(* IEC 61131-3 sources: daoli-st-library/DL_Device (part 27) *)

(* ---- FB_DL_OvenCureProfileSeq.st ---- *)
(*
  Name: FB_DL_OvenCureProfileSeq
  Category: DL_Device
  Version: 1.0.0
  Round: R89 / 2026-11-25
  开源溯源：clean-room 自研（族 涂装喷涂线，ST 开源生态实测 0 命中，无外部代码引入）
  功能：烘干炉固化温度曲线执行顺序：升温→保温→冷却→出炉许可，每段结束判据独立。
  边界条件：① 温度与速率入参全部过非有限闸（含三元素设定数组逐项），配置越域即锁故障（101）；
            ② 保温段使用独立 TON（tonSoak，PT := tSoakS），与升温/冷却段判据不同源，无双窗配比问题（R100）；
            ③ 超温判据以段 1 设定 + 15 ℃ 为上限（固化段为最高温段），越限立即锁故障（102）；
            ④ 出炉许可为单拍脉冲（内部 _bDone 置位 → 出口映射），后驻留 eDone 至启动释放；
            ⑤ 故障解除唯一路径：故障相内 xStart 释放（R152），清锁存回 eIdle。
  状态机：eIdle / eSeg1 / eSeg2 / eSeg3 / eDone / eFault（CASE 含 ELSE 兜底）。
*)
TYPE E_DL_OcpPhase :
(
    eIdle := 0,         (* 待机：等启动沿 / Idle, waiting for start edge *)
    eSeg1 := 10,        (* 段 1 升温：升到固化温度带 / Segment 1, ramp to cure band *)
    eSeg2 := 20,        (* 段 2 保温：保温窗且带内 / Segment 2, soak window in band *)
    eSeg3 := 30,        (* 段 3 冷却：冷到出炉温度 / Segment 3, cool down *)
    eDone := 40,        (* 完成相：出炉许可后驻留 / Done, holds after discharge permit *)
    eFault := 90        (* 故障相：锁存待释放 / Fault latched, awaiting release *)
);
END_TYPE

FUNCTION_BLOCK FB_DL_OvenCureProfileSeq
VAR_INPUT
    xStart : BOOL;                          (* 启动命令（上升沿起序） [-] Start command, rising edge *)
    fTempActC : REAL;                       (* 炉温实测 [℃] Oven temperature actual [degC] *)
    fTempSpC : ARRAY[1..3] OF REAL;         (* 三段温度设定（升温/保温/冷却） [℃] Segment setpoints [degC] *)
    fRampCpm : REAL;                        (* 允许升温速率 [℃/min] Allowed ramp rate [degC/min] *)
    tSoakS : TIME;                          (* 保温窗 [ms] Soak window [ms] *)
    fCoolToC : REAL;                        (* 冷却目标（出炉温度） [℃] Cool-down target [degC] *)
END_VAR
VAR_OUTPUT
    eState : E_DL_OcpPhase;                 (* 当前相 [-] Present phase *)
    nSegIdx : INT;                          (* 当前段号（0 空闲，1~3） [段] Present segment index *)
    xDone : BOOL;                           (* 出炉许可单拍脉冲 [-] Discharge permit pulse *)
    xFault : BOOL;                          (* 故障锁存标志 [-] Fault latched *)
END_VAR
VAR
    _eState : E_DL_OcpPhase := E_DL_OcpPhase.eIdle;  (* 内部相（CASE 唯一写入目标） [-] Internal phase *)
    _bDone : BOOL := FALSE;         (* 单拍完成标志（段 1 预清） [-] One-scan done flag *)
    _bFaultLatch : BOOL := FALSE;   (* 故障锁存位 [-] Fault latch *)
    _bReqFault : BOOL := FALSE;     (* 单拍故障请求（段 1 预清） [-] Fault request *)
    _bCfgBad : BOOL := FALSE;       (* 配置非法当拍量 [-] Configuration bad *)
    _nSeg : INT := 0;               (* 段号保持量 [段] Segment index hold *)
    _nErr : INT := 0;               (* 故障码锁存（101 组态 / 102 超温 / 103 非法相） [-] Latched code *)
    _nReqErr : INT := 0;            (* 当拍请求码 [-] Requested code *)
    _nI : INT := 1;                 (* 设定数组遍历索引 [-] Setpoint loop index *)
    tonSoak : TON;                  (* 保温窗（段 0 无条件调用） / Soak window timer *)
    rtStart : R_TRIG;               (* 启动沿（段 0 无条件调用） / Start edge *)
END_VAR
VAR CONSTANT
    DL_OCP_TOL : REAL := 5.0;           (* 段到位带半宽 [℃] Segment in-band half-width [degC] *)
    DL_OCP_OVER : REAL := 15.0;         (* 超温裕度 [℃] Over-temperature margin [degC] *)
    DL_OCP_T_MIN : REAL := 0.0;         (* 温度下限 [℃] Temperature floor [degC] *)
    DL_OCP_T_MAX : REAL := 400.0;       (* 温度上限 [℃] Temperature ceiling [degC] *)
    DL_OCP_R_MIN : REAL := 0.5;         (* 允许速率下限 [℃/min] Ramp rate floor [degC/min] *)
    DL_OCP_R_MAX : REAL := 50.0;        (* 允许速率上限 [℃/min] Ramp rate ceiling [degC/min] *)
    DL_OCP_SEGN : INT := 3;             (* 设定段数 [-] Segment count *)
END_VAR
(* —— 段 0：沿与保温 TON 无条件周期刷新（R7） —— *)
rtStart(CLK := xStart);                                             (* 启动沿 / Start edge *)
tonSoak(IN := (_eState = E_DL_OcpPhase.eSeg2), PT := tSoakS);       (* 保温窗 / Soak window *)
(* 非有限闸（NaN 自反 + Inf 差值自减）+ 组态域闸：标量与三元素数组全枚举（R272） *)
_bCfgBad := (fTempActC <> fTempActC) OR ((fTempActC - fTempActC) <> 0.0)
         OR (fRampCpm <> fRampCpm) OR ((fRampCpm - fRampCpm) <> 0.0)
         OR (fCoolToC <> fCoolToC) OR ((fCoolToC - fCoolToC) <> 0.0)
         OR (fTempActC < DL_OCP_T_MIN) OR (fTempActC > DL_OCP_T_MAX)
         OR (fCoolToC < DL_OCP_T_MIN) OR (fCoolToC > DL_OCP_T_MAX)
         OR (fRampCpm < DL_OCP_R_MIN) OR (fRampCpm > DL_OCP_R_MAX) OR (tSoakS <= T#0S);
FOR _nI := 1 TO DL_OCP_SEGN DO
    IF (fTempSpC[_nI] <> fTempSpC[_nI]) OR ((fTempSpC[_nI] - fTempSpC[_nI]) <> 0.0)
       OR (fTempSpC[_nI] < DL_OCP_T_MIN) OR (fTempSpC[_nI] > DL_OCP_T_MAX) THEN
        _bCfgBad := TRUE;
    END_IF
END_FOR
(* —— 段 1：单拍量预清 + 组态与超温故障请求 —— *)
_bDone := FALSE;
_bReqFault := FALSE;
_nReqErr := 0;
IF _bCfgBad THEN
    _bReqFault := TRUE; _nReqErr := 101;        (* 组态非法 / Configuration bad *)
ELSIF (NOT _bCfgBad) AND (fTempActC > (fTempSpC[1] + DL_OCP_OVER)) THEN
    _bReqFault := TRUE; _nReqErr := 102;        (* 超温 / Over-temperature *)
END_IF
(* —— 段 2：故障锁存解除（唯一路径 = 故障相内 xStart 释放，R152） —— *)
IF _bFaultLatch AND (NOT xStart) THEN
    _bFaultLatch := FALSE;                      (* 清锁存 / Clear latch *)
    _nErr := 0;                                 (* 清码 / Clear code *)
    _nSeg := 0;                                 (* 段号归零 / Segment index reset *)
    _eState := E_DL_OcpPhase.eIdle;             (* 迁回待机 / Back to idle *)
END_IF
(* —— 段 3：主状态机（ENUM + CASE，ELSE 兜底） —— *)
CASE _eState OF
E_DL_OcpPhase.eIdle:
    IF rtStart.Q AND (NOT _bFaultLatch) THEN
        _nSeg := 1;                             (* 段 1 起算 / Segment 1 begins *)
        _eState := E_DL_OcpPhase.eSeg1;
    END_IF
E_DL_OcpPhase.eSeg1:
    IF ABS(fTempActC - fTempSpC[1]) <= DL_OCP_TOL THEN
        _nSeg := 2;                             (* 进带 → 保温段 / In band, soak segment *)
        _eState := E_DL_OcpPhase.eSeg2;
    END_IF
E_DL_OcpPhase.eSeg2:
    IF tonSoak.Q AND (ABS(fTempActC - fTempSpC[2]) <= DL_OCP_TOL) THEN
        _nSeg := 3;                             (* 保温窗到且带内 → 冷却段 / Soak done, cool *)
        _eState := E_DL_OcpPhase.eSeg3;
    END_IF
E_DL_OcpPhase.eSeg3:
    IF fTempActC <= fCoolToC THEN
        _bDone := TRUE;                         (* 单拍出炉许可（段 1 预清） / One-scan permit *)
        _nSeg := 0;                             (* 段号归零 / Segment index reset *)
        _eState := E_DL_OcpPhase.eDone;
    END_IF
E_DL_OcpPhase.eDone:
    IF NOT xStart THEN
        _eState := E_DL_OcpPhase.eIdle;         (* 启动释放 → 待机 / Start released, idle *)
    END_IF
E_DL_OcpPhase.eFault:
    _nSeg := 0;                                 (* 故障相驻留：段号清零供 HMI 判别 / Residency *)
ELSE
    _bReqFault := TRUE;                         (* 非法相兜底 / Illegal phase fallback *)
    _nReqErr := 103;
END_CASE
(* —— 段 4：故障请求统一落地（唯一锁存点 + 同步迁相，R187/R252） —— *)
IF _bReqFault AND (NOT _bFaultLatch) THEN
    _bFaultLatch := TRUE;                       (* 锁存 / Latch *)
    _nErr := _nReqErr;                          (* 码锁存回放 / Latched code *)
    _eState := E_DL_OcpPhase.eFault;            (* 同步迁相 / Migrate to fault *)
END_IF
(* —— 段 5：统一出口（各出口单点赋值） —— *)
eState := _eState;
nSegIdx := _nSeg;
xDone := _bDone;
xFault := _bFaultLatch;
END_FUNCTION_BLOCK

(* ---- FB_DL_OvenDoorInterlock.st ---- *)
//==============================================================================
// 功能块：FB_DL_OvenDoorInterlock ｜ 中文名称：烘箱炉门-氮气-温区三联锁
// 所属子库：DL_Device ｜ 版本：v1.0.0 ｜ 兼容：CODESYS V3.5+ / TwinCAT 3 / 汇川 InoProShop
// 功能描述：烘箱炉门开门三联锁——门已关确认 → 氮气置换完成 → 温区温度
//           低于开门上限，三条件全满才放行开锁；任一失守立即回锁定态并
//           锁存失守原因。先置换后开门（锂电干燥环节安全前置语义）。
// 开源溯源 (Origin)：道莅 clean-room 防御性实现
// 单位表：T[°C] / 联锁条件[—]
// 错误码表：16#0003_017C 信息级（放行时温度接近上限，提示性，不置
//           bError）/ 16#0003_017D 预留禁用（不得挪用）/ 16#0003_034B
//           故障级（组态非法：开门温度上限 <= 0；或温度非有限，安全侧
//           拒绝放行，置 bError）/ 16#0003_034C 故障级（确认矛盾：门未
//           处于放行态而门关反馈消失，置 bError）/ 16#0003_034D 故障级
//           兜底（状态机落 ELSE，置 bError 并回锁定）
// 状态机：E_DL_OvenDoorState（eLocked=0 / ePurging=10 / eTempHigh=20 /
//           eReleased=30 / eFault=99），CASE 含 ELSE 兜底，ELSE 置 034D
//           并回 eLocked
// 边界行为：① 三条件任一失守 → 回 eLocked 并锁存最近失守原因码；②
//           fOpenTempMaxC <= 0 → 故障 034B 锁存（组态非法）；③ 温度非
//           有限 → 故障 034B 复用（R90）+ 拒绝放行（安全侧默认：非法值
//           绝不放行开门）；④ 温度迟滞按 FC_DL_Hysteresis 语义内联实现
//           （放行阈 <= 上限，回锁阈 > 上限 + 2 K 迟滞带）；⑤ 非放行态
//           下门关反馈消失 → 034C 故障转 eFault（未授权开门，安全侧全锁）。
// 依赖纪律：仅 Standard.library + 同库契约（无跨子库调用；温度迟滞内联，
//           依赖收窄声明：Device 不调用 DL_Base 的 FC_DL_Hysteresis，
//           迟滞语义在本件内联，改动任一侧须复核另一侧）。
// 修订历史：v1.0.0 2026-11-17 首版（R23 派单 · ROADMAP 锂电 P1 §350 + T2-8 互锁语义次源）
//==============================================================================

(*------------------------------------------------------------------------------
 * 枚举: E_DL_OvenDoorState（归属本功能块，同文件发布，全库唯一定义）
 * 含义: 炉门三联锁相位，每个成员在 CASE 中有且仅有一个标签。
 *-----------------------------------------------------------------------------*)
TYPE E_DL_OvenDoorState :
(
    eLocked   := 0,   // 锁定：门锁未放行，等开门请求与三条件 / Locked, waiting for the request and the three conditions
    ePurging  := 10,  // 置换中：门已关，等氮气置换完成确认 / Purging, door closed, waiting for the N2 purge confirmation
    eTempHigh := 20,  // 温度高：置换已完成，等温区降到开门上限以下 / Temperature high, waiting for cool-down below the limit
    eReleased := 30,  // 已放行：开锁输出有效，允许开门 / Released, unlock output active
    eFault    := 99   // 故障：组态非法/确认矛盾/非有限温度/非法状态 / Fault, illegal config, contradiction or non-finite temperature
);
END_TYPE

FUNCTION_BLOCK FB_DL_OvenDoorInterlock
VAR_INPUT
    bDoorClosedFb  : BOOL;                  // 门已关到位反馈 [—] / Door-closed feedback
    bN2PurgeOk     : BOOL;                  // 氮气置换完成 [—] / N2 purge complete
    fZoneTempC     : LREAL;                 // 温区实测温度 [摄氏度] / Measured zone temperature [degC]
    fOpenTempMaxC  : LREAL := 45.0;         // 允许开门温度上限 [摄氏度]，须 > 0 / Door-open temperature ceiling [degC], must be > 0
    bDoorOpenCmd   : BOOL;                  // 开门请求 [—]，电平有效 / Door-open request, level active
    bReset         : BOOL;                  // 故障复位 [—]，上升沿退出 eFault / Fault reset, rising edge leaves the fault state
END_VAR
VAR_OUTPUT
    bDoorUnlock    : BOOL;                  // 开锁放行 [—] / Door unlock release
    eInterlockState: E_DL_OvenDoorState;    // 联锁相位 [—] / Interlock phase
    eErr           : UDINT;                 // 错误码，0 = 无错 / Error code, 0 = no error
    bError         : BOOL;                  // 故障级标志，仅故障级错误置位 / Fault-class flag, set only on fault-level codes
    bValid         : BOOL;                  // 输出可用标志 / Outputs usable flag
END_VAR
VAR
    rtOpenReq      : R_TRIG;                // 开门请求上升沿，段 6 无条件刷新 / Open-request rising edge
    _eState        : E_DL_OvenDoorState := E_DL_OvenDoorState.eLocked; // 当前相位 / Current phase
    _bInit         : BOOL := FALSE;         // 首扫标志，初值 FALSE 取非判定 / First-scan flag, tested negated
    _bCfgBad       : BOOL;                  // 组态非法锁存 / Illegal configuration latch
    _bFiniteBad    : BOOL;                  // 温度非有限锁存 / Non-finite temperature latch
    _bIllegal      : BOOL;                  // 非法状态标志 / Illegal state flag
    _bNearLimit    : BOOL;                  // 放行时温度接近上限标志 / Near-limit flag at release
END_VAR
VAR CONSTANT
    DL_OVN_HYST    : LREAL := 2.0;          // 温度迟滞带 [K]，回锁阈 = 上限 + 迟滞 / Temperature hysteresis band [K]
    DL_OVN_NEAR    : LREAL := 5.0;          // 接近上限提示带 [K] / Near-limit notice band [K]
    DL_OVN_INF     : LREAL := 1.7976931348623157E308; // LREAL 幅值上限 / LREAL magnitude ceiling
END_VAR

(*------------------------------------------------------------------------------
 * 段 1｜每拍预置：输出先全断（安全侧），单拍标志预清零
 *      Outputs cleared first, fail-safe side, one-shot flags pre-cleared
 *-----------------------------------------------------------------------------*)
bDoorUnlock := FALSE;                       // 开锁输出先清（安全侧默认断） / Unlock preset FALSE, fail-safe
eErr        := 16#0000_0000;                // 错误码每拍重算 / Error code recomputed
bError      := FALSE;                       // 故障标志每拍重算 / Fault flag recomputed
bValid      := FALSE;                       // 可用标志每拍重算 / Usable flag recomputed
_bIllegal   := FALSE;                       // 非法状态标志预清零 / Illegal flag pre-cleared
_bNearLimit := FALSE;                       // 接近上限标志预清零 / Near-limit flag pre-cleared

(*------------------------------------------------------------------------------
 * 段 2｜首扫初始化（IF NOT bInit 范式）
 *      First-scan initialisation
 *-----------------------------------------------------------------------------*)
IF NOT _bInit THEN
    _eState  := E_DL_OvenDoorState.eLocked; // 相位锁定起步 / Phase starts locked
    _bCfgBad := FALSE;                      // 组态锁存清零 / Config latch cleared
    _bFiniteBad := FALSE;                   // 非有限锁存清零 / Non-finite latch cleared
    _bInit   := TRUE;                       // 首扫只做一次 / The first scan runs once
END_IF

(*------------------------------------------------------------------------------
 * 段 3｜组态与输入防御闸：上限 <= 0 或温度非有限 → 034B（安全侧拒绝放行）
 *      Configuration and input defense gate, fail-safe refusal
 *-----------------------------------------------------------------------------*)
IF fOpenTempMaxC <= 0.0 THEN
    _bCfgBad := TRUE;                       // 组态非法锁存 / Illegal configuration latched
END_IF
IF (fZoneTempC <> fZoneTempC) OR (ABS(fZoneTempC) > DL_OVN_INF) THEN
    _bFiniteBad := TRUE;                    // 温度非有限锁存（复用 034B，R90） / Non-finite temperature latched, code reused
END_IF
IF _bCfgBad OR _bFiniteBad THEN
    _eState := E_DL_OvenDoorState.eFault;   // 任何组态/输入异常都转故障态 / Any config or input anomaly goes to fault
END_IF

(*------------------------------------------------------------------------------
 * 段 4｜确认矛盾闸：门未处于放行态而门关反馈消失 → 未授权开门 034C
 *      Contradiction gate: door feedback lost outside the released phase
 *-----------------------------------------------------------------------------*)
IF (_eState <> E_DL_OvenDoorState.eReleased)
   AND (_eState <> E_DL_OvenDoorState.eFault) AND (NOT bDoorClosedFb) THEN
    _eState := E_DL_OvenDoorState.eFault;   // 未授权开门，转故障全锁 / Unauthorized door opening, fault with full lock
    eErr    := 16#0003_034C;                // 故障级：确认矛盾 / Fault: confirmation contradiction
    bError  := TRUE;                        // 置故障标志 / Raise the fault flag
END_IF

(*------------------------------------------------------------------------------
 * 段 5｜R_TRIG 无条件刷新（R40：CASE 之外每拍必调）
 *      R_TRIG refreshed unconditionally per R40
 *-----------------------------------------------------------------------------*)
rtOpenReq(CLK := bDoorOpenCmd);             // 开门请求上升沿 / Open-request rising edge

(*------------------------------------------------------------------------------
 * 段 6｜相位机（只做迁移；输出在段 7 按相置位）
 *      Phase machine, transitions only, outputs assigned in segment seven
 *-----------------------------------------------------------------------------*)
CASE _eState OF

    E_DL_OvenDoorState.eLocked:            // 锁定：等开门请求与氮气置换
        IF rtOpenReq.Q THEN
            IF bN2PurgeOk THEN
                _eState := E_DL_OvenDoorState.eTempHigh; // 置换已完成，直入温度评估 / Purge done, go to the temperature gate
            ELSE
                _eState := E_DL_OvenDoorState.ePurging;  // 置换未完成，先置换后开门 / Purge pending, purge first
            END_IF
        END_IF

    E_DL_OvenDoorState.ePurging:           // 置换中：等氮气置换完成
        IF bN2PurgeOk THEN
            _eState := E_DL_OvenDoorState.eTempHigh; // 置换完成，进温度评估 / Purge complete, to the temperature gate
        ELSIF NOT bDoorOpenCmd THEN
            _eState := E_DL_OvenDoorState.eLocked;   // 请求撤销，回锁定 / Request dropped, back to locked
        END_IF

    E_DL_OvenDoorState.eTempHigh:          // 温度门：降到上限以下才放行
        IF (NOT bDoorOpenCmd) THEN
            _eState := E_DL_OvenDoorState.eLocked;   // 请求撤销，回锁定 / Request dropped, back to locked
        ELSIF fZoneTempC <= fOpenTempMaxC THEN
            _eState := E_DL_OvenDoorState.eReleased; // 温度达标，放行 / Temperature within the limit, release
        END_IF

    E_DL_OvenDoorState.eReleased:          // 已放行：超迟滞带或请求撤销即回锁
        IF (fZoneTempC > fOpenTempMaxC + DL_OVN_HYST) OR (NOT bDoorOpenCmd) THEN
            _eState := E_DL_OvenDoorState.eLocked;   // 温度超迟滞带或请求撤销，回锁 / Beyond the hysteresis band or request dropped
        END_IF

    E_DL_OvenDoorState.eFault:             // 故障：原因消失且复位沿才回锁定
        IF bReset AND (NOT _bCfgBad) AND (NOT _bFiniteBad) AND bDoorClosedFb THEN
            _bCfgBad    := FALSE;          // 清组态锁存（组态引脚已修正） / Clear the config latch, the pin is fixed
            _bFiniteBad := FALSE;          // 清非有限锁存（温度已恢复） / Clear the non-finite latch
            _eState     := E_DL_OvenDoorState.eLocked; // 回锁定 / Back to locked
        END_IF

    ELSE                                   // 非法状态兜底（R21：CASE 必带 ELSE）
        _bIllegal := TRUE;                 // 标记非法状态 / Flag the illegal state
        _eState   := E_DL_OvenDoorState.eLocked; // 回锁定（安全侧） / Back to locked, fail-safe
END_CASE

(*------------------------------------------------------------------------------
 * 段 7｜输出置位与码位出口
 *      Output assignment and the code outlet
 *-----------------------------------------------------------------------------*)
IF _eState = E_DL_OvenDoorState.eReleased THEN
    bDoorUnlock := TRUE;                    // 放行态开锁输出 / Unlock output in the released phase
    IF fZoneTempC > fOpenTempMaxC - DL_OVN_NEAR THEN
        _bNearLimit := TRUE;                // 放行时温度接近上限 / Near the limit at release
    END_IF
END_IF

IF _bIllegal THEN
    eErr   := 16#0003_034D;                 // 故障级：状态机兜底 / Fault: state machine fallback
    bError := TRUE;                         // 置故障标志 / Raise the fault flag
ELSIF _bCfgBad OR _bFiniteBad THEN
    eErr   := 16#0003_034B;                 // 故障级：组态非法或温度非有限（R90 复用） / Fault: illegal config or non-finite temperature
    bError := TRUE;                         // 置故障标志 / Raise the fault flag
ELSIF (_eState = E_DL_OvenDoorState.eFault) THEN
    eErr   := 16#0003_034C;                 // 故障级：确认矛盾保持显示 / Fault: contradiction held
    bError := TRUE;                         // 置故障标志 / Raise the fault flag
ELSIF _bNearLimit THEN
    eErr := 16#0003_017C;                   // 信息级：放行时温度接近上限 / Info: near-limit release
END_IF

bValid := (NOT bError) AND (_eState <> E_DL_OvenDoorState.eFault); // 故障态输出不可用 / Outputs unusable in fault
END_FUNCTION_BLOCK

(* ---- FB_DL_PaintRobotPathSeq.st ---- *)
(*
  Name: FB_DL_PaintRobotPathSeq
  Category: DL_Device
  Version: 1.0.0
  Round: R89 / 2026-11-25
  开源溯源：clean-room 自研（族 涂装喷涂线，ST 开源生态实测 0 命中，无外部代码引入）
  功能：喷涂机器人轨迹段执行顺序（含枪距补偿）：按段完成沿推进段号，输出段号、枪距补偿量与轨迹完成脉冲。
  边界条件：① 枪距两入参过非有限闸；总段数与段索引按 1~999 域闸拦截，越域即故障（101）；
            ② 段完成沿用 R_TRIG 在段 0 无条件刷新（R7），禁放入 CASE 分支；
            ③ 枪距补偿 = 设定 − 实测，钳 ±5 mm（伺服补偿行程死区外的机械限）；
            ④ 完成脉冲两段式：相内置 _bDone，出口统一映射单拍（R187）；
            ⑤ 故障解除唯一路径：故障相内 xStart 释放（R152），清锁存回 eIdle。
  状态机：eIdle / eRun / eDone / eFault（CASE 含 ELSE 兜底）。
*)
TYPE E_DL_DpsState :
(
    eIdle  := 0,        (* 待机：等启动沿 / Idle, waiting for start edge *)
    eRun   := 10,       (* 执行相：按段完成沿推进 / Running, advancing by segment done edge *)
    eDone  := 20,       (* 完成相：保持至启动释放 / Done, holds until start released *)
    eFault := 90        (* 故障相：锁存待释放 / Fault latched, awaiting release *)
);
END_TYPE

FUNCTION_BLOCK FB_DL_PaintRobotPathSeq
VAR_INPUT
    xStart : BOOL;              (* 启动命令（上升沿起序） [-] Start command, rising edge *)
    nSegTotal : INT;            (* 轨迹总段数 [段] Total segment count *)
    nSegIdxIn : INT;            (* 起始段索引 [段] Initial segment index *)
    fGunDistActMm : REAL;       (* 枪距实测 [mm] Gun distance actual [mm] *)
    fGunDistSpMm : REAL;        (* 枪距设定 [mm] Gun distance setpoint [mm] *)
    xSegDone : BOOL;            (* 当前段完成反馈（上升沿有效） [-] Segment done feedback *)
END_VAR
VAR_OUTPUT
    nSegIdxOut : INT;           (* 当前段索引 [段] Present segment index *)
    fGunDistCompMm : REAL;      (* 枪距补偿量 [mm] Gun distance compensation [mm] *)
    xPathDone : BOOL;           (* 轨迹完成单拍脉冲 [-] One-scan path done pulse *)
    xFault : BOOL;              (* 故障锁存标志 [-] Fault latched *)
END_VAR
VAR
    _eState : E_DL_DpsState := E_DL_DpsState.eIdle;  (* 内部相（CASE 唯一写入目标） [-] Internal phase *)
    _bDone : BOOL := FALSE;         (* 单拍完成标志（段 1 预清） [-] One-scan done flag *)
    _bFaultLatch : BOOL := FALSE;   (* 故障锁存位 [-] Fault latch *)
    _bReqFault : BOOL := FALSE;     (* 单拍故障请求（段 1 预清） [-] Fault request *)
    _bCfgBad : BOOL := FALSE;       (* 配置非法当拍量 [-] Configuration bad *)
    _nSeg : INT := 1;               (* 段索引保持量 [段] Segment index hold *)
    _fComp : REAL := 0.0;           (* 枪距补偿保持量 [mm] Compensation hold [mm] *)
    rtSeg : R_TRIG;                 (* 段完成沿（段 0 无条件调用） / Segment done edge *)
    rtStart : R_TRIG;               (* 启动沿（段 0 无条件调用） / Start edge *)
END_VAR
VAR CONSTANT
    DL_DPS_COMP_MAX : REAL := 5.0;      (* 补偿量行程限 [mm] Compensation stroke limit [mm] *)
    DL_DPS_SEG_MAX : INT := 999;        (* 段数上限 [段] Segment count ceiling *)
    DL_DPS_DIST_MIN : REAL := 10.0;     (* 枪距下限 [mm] Gun distance floor [mm] *)
    DL_DPS_DIST_MAX : REAL := 400.0;    (* 枪距上限 [mm] Gun distance ceiling [mm] *)
END_VAR
(* —— 段 0：两沿无条件周期刷新（R7） —— *)
rtStart(CLK := xStart);                     (* 启动沿 / Start edge *)
rtSeg(CLK := xSegDone);                     (* 段完成沿 / Segment done edge *)
(* 非有限闸（NaN 自反 + Inf 差值自减）+ 域闸：两枪距入参与段数全枚举（R272） *)
_bCfgBad := (fGunDistActMm <> fGunDistActMm) OR ((fGunDistActMm - fGunDistActMm) <> 0.0)
         OR (fGunDistSpMm <> fGunDistSpMm) OR ((fGunDistSpMm - fGunDistSpMm) <> 0.0)
         OR (fGunDistActMm < DL_DPS_DIST_MIN) OR (fGunDistActMm > DL_DPS_DIST_MAX)
         OR (fGunDistSpMm < DL_DPS_DIST_MIN) OR (fGunDistSpMm > DL_DPS_DIST_MAX)
         OR (nSegTotal < 1) OR (nSegTotal > DL_DPS_SEG_MAX)
         OR (nSegIdxIn < 1) OR (nSegIdxIn > nSegTotal);
(* 枪距补偿：设定 − 实测，钳 ±行程限 *)
_fComp := fGunDistSpMm - fGunDistActMm;
IF _fComp > DL_DPS_COMP_MAX THEN
    _fComp := DL_DPS_COMP_MAX;
ELSIF _fComp < (0.0 - DL_DPS_COMP_MAX) THEN
    _fComp := 0.0 - DL_DPS_COMP_MAX;
END_IF
(* —— 段 1：单拍量预清 + 组态故障请求 —— *)
_bDone := FALSE;
_bReqFault := FALSE;
IF _bCfgBad THEN
    _bReqFault := TRUE;                     (* 组态非法：段数/枪距越域 / Configuration bad *)
END_IF
(* —— 段 2：故障锁存解除（唯一路径 = 故障相内 xStart 释放，R152） —— *)
IF _bFaultLatch AND (NOT xStart) THEN
    _bFaultLatch := FALSE;                  (* 清锁存 / Clear latch *)
    _nSeg := 1;                             (* 段号归位 / Segment index reset *)
    _eState := E_DL_DpsState.eIdle;         (* 迁回待机 / Back to idle *)
END_IF
(* —— 段 3：主状态机（ENUM + CASE，ELSE 兜底） —— *)
CASE _eState OF
E_DL_DpsState.eIdle:
    IF rtStart.Q AND (NOT _bFaultLatch) THEN
        _nSeg := nSegIdxIn;                 (* 按外部起始段进入 / Start from given segment *)
        _eState := E_DL_DpsState.eRun;
    END_IF
E_DL_DpsState.eRun:
    IF rtSeg.Q THEN
        IF _nSeg < nSegTotal THEN
            _nSeg := _nSeg + 1;             (* 推进一段 / Advance one segment *)
        ELSE
            _bDone := TRUE;                 (* 末段完成：单拍脉冲 / Last segment done *)
            _eState := E_DL_DpsState.eDone;
        END_IF
    END_IF
E_DL_DpsState.eDone:
    IF NOT xStart THEN
        _eState := E_DL_DpsState.eIdle;     (* 启动释放 → 待机 / Start released, idle *)
    END_IF
E_DL_DpsState.eFault:
    _fComp := fGunDistSpMm - fGunDistActMm; (* 故障相驻留：补偿量照算供追溯，不迁相 *)
ELSE
    _bReqFault := TRUE;                     (* 非法相兜底 / Illegal phase fallback *)
END_CASE
(* —— 段 4：故障请求统一落地（唯一锁存点 + 同步迁相，R187/R252） —— *)
IF _bReqFault AND (NOT _bFaultLatch) THEN
    _bFaultLatch := TRUE;                   (* 锁存 / Latch *)
    _eState := E_DL_DpsState.eFault;        (* 同步迁相 / Migrate to fault *)
END_IF
(* —— 段 5：统一出口（各出口单点赋值；补偿量在段 0 已按行程限钳定） —— *)
nSegIdxOut := _nSeg;
(* 出口非有限/越界闸：NOT(x<=lim) 对 NaN 为真，防补偿量 NaN 直穿 *)
IF NOT ((_fComp <= 1000.0) AND (_fComp >= -1000.0)) THEN
    _fComp := 0.0;                          (* 归零补偿，保持原枪距 / Zero comp, keep gun distance *)
END_IF
fGunDistCompMm := _fComp;
xPathDone := _bDone;
xFault := _bFaultLatch;
END_FUNCTION_BLOCK

(* ---- FB_DL_ParallelGripper.st ---- *)
(*
    FB_DL_ParallelGripper —— 平行夹爪实现（实现 I_DL_Gripper）
    ------------------------------------------------------------------
    分类      : DL_Device / Actuator
    前缀      : FB_DL_
    版本      : 1.0.1
    溯源      : T2-6 Rockwell AOI（只借「设备级 AOI 粒度」分类事实）；
                T1-5 开源契约-实现分离范式（仅借分层思想）；
                状态机、超时策略、空夹语义、码位 100% 自有；clean-room 重写，
                未复制任何闭源厂商源码，参考实现仅限 MIT/Apache 许可
    平台      : 纯 IEC 61131-3，CODESYS V3.5+ / TwinCAT 3 / InoProShop 通用
    作者      : 道莅代码库 · PLC编程专家（R18）
    ------------------------------------------------------------------
    功能说明  : 三段动作（驱动 → 到位确认 → 夹持力保持），含单动作超时、在位与命令
                矛盾判定、无件闭合（空夹）判定；实现 I_DL_Gripper 全部属性与方法；
                不直接写输出地址：电磁阀 / 伺服指令经 bValveOut 输出引脚由上层映射，
                换品牌只改映射层；
                安全约定：bEnable 为 FALSE、复位沿、故障态三者都在同一拍把 bValveOut
                清为 FALSE（断开驱动），绝不把「清使能」当成「保持夹持」，防夹持件掉落；
                超时参数本身非法会让超时保护失效，故 032A 同时承担「动作超时」与
                「超时参数非法」两个同源语义；
                空夹（闭合到位但无工件）是合法工况，只置信息码与 bLoadOpen，不停线。
    接口实现  : I_DL_Gripper 的七个只读属性（bOpened / bClosed / bWorkpiecePresent /
                fWidth / eHealth / uErrorId / bError）与四个方法全部在本文件尾部落地。
                五个契约量（bOpened / bClosed / bWorkpiecePresent / fWidth / bError）
                只以属性形态对外，不再另设同名输出引脚——同名成员在同一功能块命名空间
                内冲突，会出现三平台编译阻断，故按属性优先原则收敛，契约语义一字不减。
    错误码    : 16#0003_0166 空夹到位 / 开合命令同拍闭合优先 / 力给定超域已钳位——信息级，不置故障
                16#0003_0167 预留禁用（信息级，不得挪用）
                16#0003_032A 动作超时（含超时参数非法）——故障级，转故障态并断驱动
                16#0003_032B 在位信号与命令矛盾，或状态机落 ELSE 兜底——故障级，转故障态
                16#0003_032C 预留禁用（故障级，不得挪用）
    码位总账  : 16#0003_0166 用 / 16#0003_0167 预留 ｜ 16#0003_032A 用 / 16#0003_032B 用 / 16#0003_032C 预留
    状态机    : E_DL_GripperState（eIdle / eOpening / eClosing / eHolding / eFault），
                CASE 含 ELSE 兜底，兜底固定置 eFault 与 032B
    采样约定  : fbTrigReset / fbMove / fbConfirm 三个实例均在本体首部无条件调用，
                IN 引脚承载全部条件，绝不把定时器放进 IF；两个定时器分别服务超时与
                到位确认，互不干扰。
    修订记录  : 2026-11-16 v1.0.0 首次入库（R18）
                2026-11-16 v1.0.1 R18 终审修复：METHOD Close 的形参 fForceSetpoint 原先只登记请求、未落到
                力通道，被同名引脚给定静默覆盖（接口承诺「按指定夹持力闭合」实际不生效）；新增方法力锁存
                fForceMeth / bForceMeth，段 4 改为方法优先、用后即清，复位路径一并清理。对外引脚与属性零变更。
*)

(*-----------------------------------------------------------------------------
 * 枚举: E_DL_GripperState（归属本实现块，与其同文件发布）
 * 含义: 平行夹爪动作状态机离散态，步长 10 留空位，故障态取 99 排末位
 *----------------------------------------------------------------------------*)
TYPE E_DL_GripperState :
(
    eIdle    := 0,     // 空闲：无动作，驱动断开 / Idle, no motion, drive released
    eOpening := 10,    // 张开中：等待全开到位 / Opening, waiting for the open feedback
    eClosing := 20,    // 闭合中：等待闭合到位 / Closing, waiting for the close feedback
    eHolding := 30,    // 夹持保持：闭合到位后维持夹持力 / Holding, keeps the clamping force after arrival
    eFault   := 99     // 故障锁存：超时 / 矛盾 / 非法状态，仅复位清除 / Fault latched, timeout, conflict or illegal state, reset only
) UINT;
END_TYPE

FUNCTION_BLOCK FB_DL_ParallelGripper IMPLEMENTS I_DL_Gripper
VAR_INPUT
    bEnable            : BOOL;                 // 使能，FALSE 撤所有输出并回空闲 / enable, FALSE drops every output and returns to idle
    bReset             : BOOL;                 // 复位，上升沿清故障 / reset, rising edge clears the fault
    bCmdOpen           : BOOL;                 // 张开请求，与闭合同拍时闭合优先 / open request, the close request wins when both are set
    bCmdClose          : BOOL;                 // 闭合请求 / close request
    fForceSetpoint     : REAL := 50.0;         // 夹持力给定 [%]，范围 0.0~100.0，超域钳位 / clamping force setpoint [%], range 0.0~100.0, clamped outside
    bOpenFeedback      : BOOL;                 // 全开到位传感器 / fully open position sensor
    bCloseFeedback     : BOOL;                 // 闭合到位传感器 / fully closed position sensor
    bWorkpieceFeedback : BOOL;                 // 工件在位传感器 / workpiece present sensor
    tMoveTime          : TIME := T#2S;         // 单动作超时 [ms]，范围 100~10000 / single action timeout [ms], range 100~10000
    tConfirmTime       : TIME := T#100MS;      // 到位确认时间 [ms]，范围 0~1000 / arrival confirmation time [ms], range 0~1000
END_VAR
VAR_OUTPUT
    bValveOut         : BOOL;                  // 驱动输出，TRUE 为闭合方向，由上层映射到物理点 / drive output, TRUE closes, mapped to the physical point upstream
    fForceOut         : REAL;                  // 实际下发夹持力，钳位后 [%] / clamping force actually issued after clamping [%]
    bBusy             : BOOL;                  // 动作中 / action in progress
    bDone             : BOOL;                  // 到位单周期脉冲 / arrival single-cycle pulse
    tElapsed          : TIME;                  // 本动作已耗时 [ms] / elapsed time of the current action [ms]
    eErr              : UDINT;                 // 错误码，0=正常 / error id, 0=ok
    bLoadOpen         : BOOL;                  // 空夹（闭合到位但无工件）/ empty clamp, closed without a workpiece
END_VAR
VAR
    fbTrigReset  : R_TRIG;                     // 复位沿检测实例，本体首部无条件刷新 / reset edge instance, refreshed unconditionally
    fbMove       : TON;                        // 单动作超时定时器，本体首部无条件刷新 / action timeout timer, refreshed unconditionally
    fbConfirm    : TON;                        // 到位确认定时器，本体首部无条件刷新 / arrival confirmation timer, refreshed unconditionally
    eState       : E_DL_GripperState := E_DL_GripperState.eIdle; // 内部状态机步序 / internal state machine step
    bPendOpen    : BOOL;                       // 方法张开请求锁存，由主体消费 / method open request latch, consumed by the body
    bPendClose   : BOOL;                       // 方法闭合请求锁存 / method close request latch
    bPendRelease : BOOL;                       // 方法泄力请求锁存 / method release request latch
    bPendClear   : BOOL;                       // 方法清故障请求锁存 / method clear fault request latch
    fForceEff    : REAL;                       // 生效夹持力，钳位后 [%] / effective clamping force after clamping [%]
    bAtTarget    : BOOL;                       // 本拍到位反馈成立标志 / arrival feedback valid this cycle
    bFaultLatch  : BOOL;                       // 故障锁存位，仅复位或方法复位清除 / fault latch, cleared by reset or the method only
    bLoadLatch   : BOOL;                       // 空夹锁存，复位清除 / empty clamp latch, cleared by reset
    bBothCmd     : BOOL;                       // 开合命令同拍标志 / both commands active flag
    fForceMeth   : REAL;                       // 方法给定的夹持力锁存，Close() 写入 [%] / clamping force latched by the Close method [%]
    bForceMeth   : BOOL;                       // 方法给定有效标志，段 4 消费后清 / method force valid flag, cleared after segment four consumes it
    fForceRaw    : REAL;                       // 本拍生效的原始力给定（方法优先于引脚）[%] / raw force actually in effect this cycle, the method wins over the pin [%]
END_VAR
VAR CONSTANT
    DL_GRP_FORCE_MAX  : REAL := 100.0;         // 夹持力上限 [%] / clamping force upper bound [%]
    DL_GRP_FORCE_MIN  : REAL := 0.0;           // 夹持力下限 [%] / clamping force lower bound [%]
    DL_GRP_MOVE_MIN   : TIME := T#100MS;       // 超时下限 [ms] / timeout lower bound [ms]
    DL_GRP_MOVE_MAX   : TIME := T#10S;         // 超时上限 [ms] / timeout upper bound [ms]
    DL_GRP_WIDTH_NONE : REAL := 0.0;           // 无模拟量反馈时的宽度缺省值 [mm] / default width without an analogue feedback [mm]
    DL_FLOAT_EPS      : REAL := 1.0E-6;        // 浮点判等容差 [%] / float equality tolerance [%]
END_VAR

METHOD Open : BOOL
VAR_INPUT
END_VAR
IF bFaultLatch OR (eState = E_DL_GripperState.eFault) THEN
    Open := FALSE;                             // 故障态拒绝 / rejected in the fault state
    bPendOpen := FALSE;                        // 清残留请求 / clear the stale request
ELSE
    bPendOpen := TRUE;                         // 登记张开请求，主体状态机消费 / register the request, consumed by the body
    bPendClose := FALSE;                       // 互斥注销闭合请求 / cancel the opposite request
    Open := TRUE;                              // 受理成功 / accepted
END_IF

(*-----------------------------------------------------------------------------
 * 方法: Close —— 请求闭合到指定夹持力。故障锁存期拒绝并返回 FALSE。
 *      Method Close - request closing at the given force, rejected while a fault is latched.
 *----------------------------------------------------------------------------*)
    END_METHOD

METHOD Close : BOOL
VAR_INPUT
    fForceSetpoint : REAL;                     // 目标夹持力 [%]，范围 0.0~100.0 / target clamping force [%], range 0.0~100.0
END_VAR
IF bFaultLatch OR (eState = E_DL_GripperState.eFault) THEN
    Close := FALSE;                            // 故障态拒绝 / rejected in the fault state
    bPendClose := FALSE;                       // 清残留请求 / clear the stale request
ELSE
    bPendClose := TRUE;                        // 登记闭合请求 / register the close request
    fForceMeth := fForceSetpoint;              // 锁存方法形参，由段 4 消费 / latch the method parameter, consumed by segment four
    bForceMeth := TRUE;                        // 置方法给定有效 / mark the method setpoint valid
    bPendOpen := FALSE;                        // 互斥注销张开请求 / cancel the opposite request
    Close := TRUE;                             // 受理成功 / accepted
END_IF

(*-----------------------------------------------------------------------------
 * 方法: Release —— 松开并撤力。与 Open 的区别是不驱动到位，只泄力。
 *      Method Release - drop the force without driving to the open end.
 *----------------------------------------------------------------------------*)
    END_METHOD

METHOD Release : BOOL
VAR_INPUT
END_VAR
IF bFaultLatch OR (eState = E_DL_GripperState.eFault) THEN
    Release := FALSE;                          // 故障态拒绝 / rejected in the fault state
ELSE
    bPendRelease := TRUE;                      // 登记泄力请求 / register the release request
    bPendOpen := FALSE;                        // 撤销张开请求 / cancel the open request
    bPendClose := FALSE;                       // 撤销闭合请求 / cancel the close request
    Release := TRUE;                           // 受理成功 / accepted
END_IF

(*-----------------------------------------------------------------------------
 * 方法: ClearFault —— 清故障锁存（热复位）。绝不隐式产生动作。
 *      Method ClearFault - clear the fault latch, never produces any motion.
 *----------------------------------------------------------------------------*)
    END_METHOD

METHOD ClearFault : BOOL
VAR_INPUT
END_VAR
IF bFaultLatch OR (eState = E_DL_GripperState.eFault) THEN
    bPendClear := TRUE;                        // 登记清故障请求，主体状态机消化 / register the request, consumed by the body
    ClearFault := TRUE;                        // 可复位 / resettable
ELSE
    ClearFault := FALSE;                       // 无故障可复位 / nothing to clear
END_IF

(*-----------------------------------------------------------------------------
 * 属性: bOpened（GET）—— 全开到位只读视图 / property bOpened (GET), read-only view
 *----------------------------------------------------------------------------*)
    END_METHOD

// 段 1｜边沿与两个定时器无条件周期刷新（红线：严禁放入条件分支）/ segment 1, unconditional refresh of the edge and both timers
fbTrigReset(CLK := bReset);
fbMove(IN := bEnable AND ((eState = E_DL_GripperState.eOpening) OR (eState = E_DL_GripperState.eClosing)), PT := tMoveTime); // 超时只服务动作态 / the timeout only serves the moving states
bAtTarget := ((eState = E_DL_GripperState.eOpening) AND bOpenFeedback)
          OR ((eState = E_DL_GripperState.eClosing) AND bCloseFeedback); // 到位判据按当前动作取对应反馈 / the arrival criterion picks the feedback of the current action
fbConfirm(IN := bEnable AND bAtTarget, PT := tConfirmTime); // 到位确认定时器 / arrival confirmation timer

// 段 2｜输出与错误状态预置 / segment 2, preset outputs and error status
bDone := FALSE;                                // 到位脉冲先清 / clear the arrival pulse first
eErr := 0;                                     // 预置无错误 / preset no error
bBusy := FALSE;                                // 预置不忙 / preset not busy
bValveOut := FALSE;                            // 驱动先按断开预置，安全侧 / preset the drive released, safe side
fForceOut := DL_GRP_FORCE_MIN;                 // 力输出先归零 / force output to zero first

// 段 3｜超时参数闸：参数非法会让超时保护失效，与动作超时同码 / segment 3, timeout parameter gate
IF (tMoveTime < DL_GRP_MOVE_MIN) OR (tMoveTime > DL_GRP_MOVE_MAX) THEN
    eErr := 16#0003_032A;                      // 超时参数非法故障码 / illegal timeout parameter fault id
    bFaultLatch := TRUE;                       // 锁存 / latch it
    eState := E_DL_GripperState.eFault;        // 转故障态 / enter the fault state
END_IF

// 段 4｜夹持力闸：方法给定优先于引脚给定，超域钳位并置信息码 / segment 4, the method force wins over the pin, then clamp and hint
fForceRaw := fForceSetpoint;                   // 默认取引脚给定 / default to the pin setpoint
IF bForceMeth THEN
    fForceRaw := fForceMeth;                   // 方法给定优先，Close() 的形参绝不静默丢弃 / the method setpoint wins, the Close parameter is never silently dropped
    bForceMeth := FALSE;                       // 用后即清，绝不跨拍残留 / consumed and cleared, never leaks to the next cycle
END_IF
fForceEff := MIN(MAX(fForceRaw, DL_GRP_FORCE_MIN), DL_GRP_FORCE_MAX); // 双侧钳位 / clamp both sides
IF ABS(fForceEff - fForceRaw) > DL_FLOAT_EPS THEN
    eErr := 16#0003_0166;                      // 力给定钳位提示（信息级不置故障）/ force clamp hint, info level never raises a fault
END_IF

// 段 5｜开合同拍判定：闭合优先（安全侧）/ segment 5, simultaneous command arbitration, close wins
bBothCmd := bCmdOpen AND bCmdClose;            // 同拍判定 / simultaneous detection
IF bBothCmd THEN
    eErr := 16#0003_0166;                      // 同拍提示（信息级不置故障）/ simultaneous hint, info level never raises a fault
END_IF

// 段 6｜复位沿与清故障方法：同拍优先于动作 / segment 6, reset edge and clear fault method take priority
IF fbTrigReset.Q OR bPendClear THEN
    bFaultLatch := FALSE;                      // 清故障锁存 / clear the fault latch
    bLoadLatch := FALSE;                       // 清空夹锁存 / clear the empty clamp latch
    bPendClear := FALSE;                       // 用后即清 / consumed and cleared
    bPendOpen := FALSE;                        // 清残留请求 / clear the stale requests
    bPendClose := FALSE;                       // 清残留请求 / clear the stale requests
    bPendRelease := FALSE;                     // 清残留请求 / clear the stale requests
    bForceMeth := FALSE;                       // 清方法力给定，防复位后误用旧值 / clear the method force so a stale value cannot be reused after a reset
    eState := E_DL_GripperState.eIdle;         // 回空闲态 / back to idle
END_IF

// 段 7｜使能闸：撤所有输出并回空闲（防夹持件掉落）/ segment 7, enable gate drops every output
IF NOT bEnable THEN
    bValveOut := FALSE;                        // 驱动断开 / drive released
    fForceOut := DL_GRP_FORCE_MIN;             // 力撤除 / force removed
    bBusy := FALSE;                            // 不忙 / not busy
    bPendOpen := FALSE;                        // 清请求 / clear the requests
    bPendClose := FALSE;                       // 清请求 / clear the requests
    bPendRelease := FALSE;                     // 清请求 / clear the requests
    eState := E_DL_GripperState.eIdle;         // 回空闲 / back to idle
    tElapsed := fbMove.ET;                     // 耗时镜像 / elapsed mirror
    RETURN;                                    // 失能即出口 / disabled is the exit
END_IF

// 段 8｜动作超时：定时器到期即故障并断驱动 / segment 8, action timeout
IF fbMove.Q THEN
    eErr := 16#0003_032A;                      // 动作超时故障码 / action timeout fault id
    bFaultLatch := TRUE;                       // 锁存 / latch it
    eState := E_DL_GripperState.eFault;        // 转故障态 / enter the fault state
END_IF

// 段 9｜在位与命令矛盾判定：闭合指令已撤但闭合反馈仍在且无工件 / segment 9, presence and command conflict
IF bCloseFeedback AND (NOT bWorkpieceFeedback) THEN
    bLoadLatch := TRUE;                        // 空夹锁存（合法工况，不停线）/ latch the empty clamp, a legal condition, no line stop
    eErr := 16#0003_0166;                      // 空夹提示（信息级不置故障）/ empty clamp hint, info level never raises a fault
END_IF

// 段 10｜状态机主体（CASE 必含 ELSE 兜底，红线）/ segment 10, state machine body
CASE eState OF
    E_DL_GripperState.eIdle :
        bValveOut := FALSE;                    // 空闲断驱动 / the idle state releases the drive
        fForceOut := DL_GRP_FORCE_MIN;         // 力撤除 / force removed
        IF bPendRelease THEN
            bPendRelease := FALSE;             // 泄力请求只清标志，不产生动作 / a release request only clears its flag, no motion
        ELSIF bCmdClose OR bPendClose THEN
            bPendClose := FALSE;               // 用后即清 / consumed and cleared
            eState := E_DL_GripperState.eClosing; // 闭合优先（含同拍情形）/ close wins, including the simultaneous case
        ELSIF bCmdOpen OR bPendOpen THEN
            bPendOpen := FALSE;                // 用后即清 / consumed and cleared
            eState := E_DL_GripperState.eOpening; // 进张开态 / enter the opening state
        END_IF
    E_DL_GripperState.eOpening :
        bValveOut := FALSE;                    // 张开方向驱动 / drive in the opening direction
        fForceOut := DL_GRP_FORCE_MIN;         // 张开不加力 / no force while opening
        bBusy := TRUE;                         // 动作中 / in motion
        IF fbConfirm.Q THEN
            bDone := TRUE;                     // 到位单拍脉冲 / arrival single-cycle pulse
            bBusy := FALSE;                    // 到位不忙 / no longer busy
            eState := E_DL_GripperState.eIdle; // 张开到位回空闲 / back to idle after opening
        END_IF
    E_DL_GripperState.eClosing :
        bValveOut := TRUE;                     // 闭合方向驱动 / drive in the closing direction
        fForceOut := fForceEff;                // 下发钳位后的夹持力 / issue the clamped force
        bBusy := TRUE;                         // 动作中 / in motion
        IF fbConfirm.Q THEN
            bDone := TRUE;                     // 到位单拍脉冲 / arrival single-cycle pulse
            bBusy := FALSE;                    // 到位不忙 / no longer busy
            eState := E_DL_GripperState.eHolding; // 进夹持保持态 / enter the holding state
        END_IF
    E_DL_GripperState.eHolding :
        bValveOut := TRUE;                     // 保持夹持 / keep clamping
        fForceOut := fForceEff;                // 保持钳位后的夹持力 / keep the clamped force
        bBusy := FALSE;                        // 保持态不算动作中 / holding is not an action
        IF (NOT bCmdClose) AND (NOT bPendClose) THEN
            eState := E_DL_GripperState.eIdle; // 命令撤销即回空闲 / back to idle when the command is withdrawn
        END_IF
    E_DL_GripperState.eFault :
        bValveOut := FALSE;                    // 故障态断驱动 / the fault state releases the drive
        fForceOut := DL_GRP_FORCE_MIN;         // 力撤除 / force removed
        bBusy := FALSE;                        // 不忙 / not busy
ELSE
    eState := E_DL_GripperState.eFault;        // 非法状态一律回安全故障态 / any illegal state falls back to the safe fault state
    eErr := 16#0003_032B;                      // 兜底故障码 / fallback fault id
    bFaultLatch := TRUE;                       // 锁存 / latch it
    bValveOut := FALSE;                        // 断驱动 / release the drive
    fForceOut := DL_GRP_FORCE_MIN;             // 力撤除 / force removed
END_CASE

// 段 11｜故障锁存对外输出与属性镜像 / segment 11, fault latch output and property mirrors
bLoadOpen := bLoadLatch;                       // 空夹输出镜像 / empty clamp mirror
tElapsed := fbMove.ET;                         // 本动作已耗时 / elapsed time of the current action

(*-----------------------------------------------------------------------------
 * 方法: Open —— 请求张开。故障锁存期拒绝并返回 FALSE。
 *      Method Open - request opening, rejected with FALSE while a fault is latched.
 *----------------------------------------------------------------------------*)

PROPERTY bOpened : BOOL
bOpened := bOpenFeedback;                      // 返回全开到位反馈 / return the open position feedback

(*-----------------------------------------------------------------------------
 * 属性: bClosed（GET）—— 闭合到位只读视图 / property bClosed (GET), read-only view
 *----------------------------------------------------------------------------*)
PROPERTY bClosed : BOOL
bClosed := bCloseFeedback;                     // 返回闭合到位反馈 / return the close position feedback

(*-----------------------------------------------------------------------------
 * 属性: bWorkpiecePresent（GET）—— 工件在位只读视图 / property bWorkpiecePresent (GET)
 *----------------------------------------------------------------------------*)
PROPERTY bWorkpiecePresent : BOOL
bWorkpiecePresent := bWorkpieceFeedback;       // 返回工件在位反馈 / return the workpiece feedback

(*-----------------------------------------------------------------------------
 * 属性: fWidth（GET）—— 开口宽度只读视图（本实现不做模拟量换算）/ property fWidth (GET)
 *----------------------------------------------------------------------------*)
PROPERTY fWidth : REAL
fWidth := DL_GRP_WIDTH_NONE;                   // 无模拟量反馈时的缺省宽度 / default width without an analogue feedback

(*-----------------------------------------------------------------------------
 * 属性: eHealth（GET）—— 健康状态，引用库内唯一属主枚举 / property eHealth (GET)
 *----------------------------------------------------------------------------*)
PROPERTY eHealth : E_DL_Ne107Status
IF bFaultLatch OR (eState = E_DL_GripperState.eFault) THEN
    eHealth := E_DL_Ne107Status.eFailure;      // 有锁存故障即失败级 / a latched fault maps to the failure class
ELSE
    eHealth := E_DL_Ne107Status.eOk;           // 否则健康 / otherwise healthy
END_IF

(*-----------------------------------------------------------------------------
 * 属性: uErrorId（GET）—— 末次故障码只读视图 / property uErrorId (GET)
 *----------------------------------------------------------------------------*)
PROPERTY uErrorId : UDINT
uErrorId := eErr;                              // 返回末次错误码 / return the last error id

(*-----------------------------------------------------------------------------
 * 属性: bError（GET）—— 故障锁存只读视图 / property bError (GET)
 *----------------------------------------------------------------------------*)
PROPERTY bError : BOOL
bError := bFaultLatch OR (eState = E_DL_GripperState.eFault); // 派生式排除信息级码 / derived form excluding info-level codes
END_FUNCTION_BLOCK

(* ---- FB_DL_PhaseLossGuard.st ---- *)
(*
  ==================================================================
  组件名 Component  : FB_DL_PhaseLossGuard
  分类   Category   : DL_Device
  前缀   Naming     : FB_DL_ ｜ b/n/u/f/t/e/st 类型前缀制（R265）
  复杂度 Complexity  : 中
  版本   Version    : 1.0.0
  功能   Purpose    : 三相缺相/逆相序检测（幅差判据 + 逆相序独立码）。
  来源   Source     : self-std（三相监测公开工程语义自研）
  平台   Platform   : 纯 IEC 61131-3（比较 / ABS / R_TRIG），三平台通用
  分工声明 Split     : 与 FB_DL_PhaseNeutralImbalance 分工——后者做相零不平衡
                      统计；本件做缺相保护与逆相序判定（R216 双向互引）。
  作者   Author     : 道莅代码库 · PLC 编程专家（R61）
  归属 Ownership     : 本件无 TYPE 声明；引用件类型全部 IEC 标准原生。
  ------------------------------------------------------------------
  边界 Boundary     :
                      一 幅差判据阈值 fImbPct 提级为输入引脚并带单位 [%]（R 红线 7），
                         阈值 ≤ 0 或非有限判组态非法锁存（0706）；
                      二 非有限闸逐个点名三个电压浮点入参（R272 全量：fUA / fUB /
                         fUC），命中判缺相成因独立锁存（0704，R190 归因唯一）；
                      三 仅全相有压时才判序（防欠压误报，边界口径）：缺相或欠压
                         态不判逆相序；逆相序独立码 0705（R190 独立成员独立码）；
                      四 双锁存独立解除：bReset 上升沿清双侧锁存（恒可达，R152）；
                      五 无全局、无外部变量、无物理地址。
  错误码   Codes    :
    16#0003_0704【故障级】缺相（幅差超阈或电压非有限），锁存至复位沿
    16#0003_0705【故障级】逆相序（相序反馈为反且全相有压），锁存至复位沿
    16#0003_0706【故障级】组态非法（阈值 ≤ 0 或非有限），锁存至复位沿
  验收   Acceptance :
    算法已证（脚本）：未跑 ｜ 编译器已证（三平台）：未跑
    V1 三相 230/230/230、阈 10% → 无故障
    V2 C 相掉至 0（幅差 100%）→ 码 0704、bPhaseLoss 锁存
    V3 全相有压 + 相序反馈反 → 码 0705、bSeqReverse 锁存
  修订记录 Revision  :
    2026-11-21  v1.0.0  R61 首版（批 3 · 序号 12）
  ==================================================================
*)
FUNCTION_BLOCK FB_DL_PhaseLossGuard
VAR_INPUT
    bEnable : BOOL := TRUE;   // 使能，FALSE 时冻结判据出口（R191 声明行）/ the enable, false freezes the judgement outlet
    bReset  : BOOL := FALSE;  // 故障复位电平，上升沿清锁存 / the fault reset level
    bSeqOk  : BOOL := TRUE;   // 相序继电器反馈：TRUE 正序 / the phase sequence relay feedback
    fUA     : LREAL := 230.0; // A 相电压有效值 [伏] / the phase A voltage
    fUB     : LREAL := 230.0; // B 相电压有效值 [伏] / the phase B voltage
    fUC     : LREAL := 230.0; // C 相电压有效值 [伏] / the phase C voltage
    fImbPct : LREAL := 10.0;  // 幅差判据阈值 [%]，必须 > 0 / the unbalance threshold in percent, must be positive
END_VAR
VAR_OUTPUT
    bPhaseLoss  : BOOL := FALSE;          // 缺相锁存指示 [-] / the phase loss latched indicator
    bSeqReverse : BOOL := FALSE;          // 逆相序锁存指示 [-] / the reverse sequence latched indicator
    bError      : BOOL := FALSE;          // 故障锁存位（与锁存同源，R191）/ the fault bit from the latch
    bValid      : BOOL := FALSE;          // 判据可用标志（无故障且无组态非法）[-] / the judgement usable flag
    eErr        : UDINT := 16#0000_0000;  // 错误码，0 = 正常 / the error code, zero is ok
END_VAR
VAR
    _bInit    : BOOL := FALSE; // 首拍初始化标志（R310）/ the first scan flag
    _bLoss    : BOOL := FALSE; // 缺相锁存副本（仅复位沿清除）/ the loss latch copy
    _bRev     : BOOL := FALSE; // 逆相序锁存副本 / the reverse latch copy
    _bCfgBad  : BOOL := FALSE; // 组态非法锁存副本 / the configuration latch copy
    _bFin     : BOOL := FALSE; // 电压非有限标记（逐拍重算）/ the voltage finiteness flag recomputed
    _fMean    : LREAL := 0.0;  // 三相电压均值 [伏] / the three phase mean voltage
    _fDev     : LREAL := 0.0;  // 当前相幅差 [%] / the current phase deviation in percent
    _bAllUp   : BOOL := FALSE; // 全相有压标记（均值 > 容差）[-] / the all phases powered flag
    rtReset   : R_TRIG; // 复位沿实例，段 0 无条件刷新 / the reset edge instance
END_VAR
VAR CONSTANT
    DL_PLG_TOL : LREAL := 1.0E-6; // 全相有压均值容差 [伏] / the mean voltage tolerance
END_VAR

// 段 0｜复位沿无条件周期刷新（禁入分支，R7）/ segment 0, the unconditional refresh
rtReset(CLK := bReset); // 复位沿 / the reset edge

// 段 1｜首拍初始化与复位沿作用域（R310 / R311）/ segment 1, the first scan init and the reset scope
IF NOT _bInit THEN // 首拍一拍 / the first scan
    _bInit := TRUE; // 置首拍标志 / raise the first scan flag
    _bLoss := FALSE; // 缺相锁存显式清零 / clear the loss latch explicitly
    _bRev := FALSE; // 逆相序锁存显式清零 / clear the reverse latch explicitly
    _bCfgBad := FALSE; // 组态锁存显式清零 / clear the configuration latch explicitly
END_IF
IF rtReset.Q THEN // 复位沿（作用域：清三锁存，R311 声明）/ the reset edge with the declared scope
    _bLoss := FALSE; // 清缺相锁存（解除路径：复位沿恒可达，R152 自证）/ clear the loss latch
    _bRev := FALSE; // 清逆相序锁存 / clear the reverse latch
    _bCfgBad := FALSE; // 清组态锁存 / clear the configuration latch
END_IF

// 段 2｜组态闸与电压非有限闸（R272 全量点名，边界一二）/ segment 2, the configuration and the voltage gates
_bFin := (fUA = fUA) AND ((fUA - fUA) = (fUA - fUA))
AND (fUB = fUB) AND ((fUB - fUB) = (fUB - fUB))
AND (fUC = fUC) AND ((fUC - fUC) = (fUC - fUC)); // 三相电压逐个自反 + 差值判 / the three voltages tested term by term
IF (fImbPct <= 0.0) OR (fImbPct <> fImbPct) OR ((fImbPct - fImbPct) <> (fImbPct - fImbPct)) THEN // 阈值非法（边界一）/ an illegal threshold
    _bCfgBad := TRUE; // 锁存组态非法（0706）/ latch the configuration fault
END_IF
IF NOT _bFin THEN // 电压非有限按缺相成因独立锁存（R190 归因唯一，边界二）/ a non finite voltage latches the loss cause
    _bLoss := TRUE; // 锁存缺相（0704）/ latch the phase loss
END_IF

// 段 3｜幅差判据（电压有限且组态合法时执行，除零防护）/ segment 3, the unbalance criterion with the division guards
IF _bFin AND (NOT _bCfgBad) THEN // 判据执行前置 / the criterion preconditions
    _fMean := (fUA + fUB + fUC) / 3.0; // 三相均值（除子常量 3.0，无除零风险）/ the mean with the constant divisor
    IF ABS(_fMean) > DL_PLG_TOL THEN // 均值非零才判幅差（除零防护）/ the deviation judged on a nonzero mean
        IF (ABS(fUA - _fMean) / ABS(_fMean) * 100.0 > fImbPct)
        OR (ABS(fUB - _fMean) / ABS(_fMean) * 100.0 > fImbPct)
        OR (ABS(fUC - _fMean) / ABS(_fMean) * 100.0 > fImbPct) THEN // 任一相幅差超阈（除子已证 > 容差）/ any phase over the threshold
            _bLoss := TRUE; // 锁存缺相（0704）/ latch the phase loss
        END_IF
    ELSE // 全相零压：按缺相成因处理（判据退化安全侧）/ the all zero phases latches the loss too
        _bLoss := TRUE; // 锁存缺相 / latch the phase loss
    END_IF
    _bAllUp := ABS(_fMean) > DL_PLG_TOL; // 全相有压标记（判序前置，边界三）/ the all powered flag ahead of the sequence test
END_IF

// 段 4｜逆相序判据（仅全相有压且未缺相未组态非法时判，边界三）/ segment 4, the reverse sequence criterion with the preconditions
IF _bAllUp AND (NOT _bLoss) AND (NOT _bCfgBad) AND (NOT bSeqOk) THEN // 判序前置齐全 / the sequence preconditions met
    _bRev := TRUE; // 锁存逆相序（0705，独立成因独立码，R190）/ latch the reverse sequence
END_IF

// 段 5｜统一出口（锁存同源映射；失能冻结判据出口保持锁存值，R191）/ segment 5, the unified outlet
bPhaseLoss := _bLoss; // 缺相出口 / the loss outlet
bSeqReverse := _bRev; // 逆相序出口 / the reverse outlet
bError := _bLoss OR _bRev OR _bCfgBad; // 故障位出口 / the fault bit outlet
bValid := (NOT _bLoss) AND (NOT _bRev) AND (NOT _bCfgBad) AND bEnable; // 判据可用标志 / the usable flag
IF _bCfgBad THEN // 组态成因回放优先 / the configuration cause replays first
    eErr := 16#0003_0706; // 故障级：阈值组态非法 / fault grade, the illegal threshold
ELSIF _bLoss THEN // 缺相成因 / the loss cause
    eErr := 16#0003_0704; // 故障级：缺相锁存回放 / fault grade, the phase loss replayed
ELSIF _bRev THEN // 逆相序成因 / the reverse cause
    eErr := 16#0003_0705; // 故障级：逆相序锁存回放 / fault grade, the reverse sequence replayed
ELSE // 无故障 / no fault
    eErr := 16#0000_0000; // 正常 / ok
END_IF
END_FUNCTION_BLOCK

(* ---- FB_DL_PhaseNeutralImbalance.st ---- *)
(*
  FB_DL_PhaseNeutralImbalance  —  三相不平衡度与中性线电流判据 / Three-phase imbalance and neutral current criterion
  分类 Category : DL_Device
  码位 Code     : 16#03_2_03
  版本 Version  : 1.0.0
  溯源 Source   : NAMUR NE107 语义借鉴 · clean-room 实现，仅借分类/参数域/命名，未复制源码
  功能 Function : 1) 三相电压/电流任一为 0 或 NaN 时改判「缺相」，不计算不平衡率（除零前置）；
                  2) 不平衡率按「最大相偏差 / 三相均值 × 100%」定义（见下方定义段），分警告/跳闸两级；
                  3) 中性线电流超限与不平衡分级各自独立码值（归因唯一，不合并）。
  边界 Boundary : ① 三相任一为 0 或 NaN 改判缺相（除零前置），不出不平衡率；
                  ② 不平衡率定义在头注释写死（最大相偏差 / 均值）；
                  ③ 中性线超限与不平衡分级各自独立码值；
                  ④ 输出三行同向：不平衡率 → 分级标志 → 缺相标志。
  依赖 Depends  : None

  不平衡率定义（写死，不随组态变化）:
    fImbalPct = MAX(|Vi − Vavg|) / Vavg × 100%，Vi 为三线电压，Vavg 为三线均值 [V]。
    电流不平衡同式，本件对电压与电流分别计算后取较大者作为综合不平衡率。
  码表 Error codes（本件子码步进 16#10，避让邻件码位）:
    16#0002_0303 故障级：不平衡跳闸级越限（保持型，需 bReset）
    16#0002_0313 故障级：中性线电流越限（独立码，需 bReset）
    16#0002_0323 信息级：缺相识别（不置 bError，由上层停机逻辑处理）
*)

TYPE E_DL_PniPhase :
(
    eIdle    := 0,   // 空闲 / Idle
    eMeasure := 10,  // 测量判定 / Measurement
    eWarn    := 20,  // 不平衡警告 / Imbalance warning
    eTrip    := 30,  // 不平衡跳闸 / Imbalance trip
    eLoss    := 40,  // 缺相 / Phase loss
    eFault   := 90   // 故障锁定 / Fault locked
);
END_TYPE

FUNCTION_BLOCK FB_DL_PhaseNeutralImbalance
VAR_INPUT
    bEnable      : BOOL;                          // 总使能，FALSE 回空闲 / Master enable
    bReset       : BOOL;                          // 复位，上升沿清跳闸与中性线锁存 / Reset
    afVoltV      : ARRAY[1..3] OF REAL;           // 三线电压 [V]，域 0~600 / Line voltages [V]
    afCurrA      : ARRAY[1..3] OF REAL;           // 三线电流 [A]，域 0~2000 / Line currents [A]
    fNeutralA    : REAL;                          // 中性线电流 [A]，域 0~2000 / Neutral current [A]
    fImbalWarnPct: REAL := 10.0;                  // 不平衡警告门限 [%]，域 > 0 / Imbalance warning limit [%]
    fImbalTripPct: REAL := 20.0;                  // 不平衡跳闸门限 [%]，须 > 警告门限 / Imbalance trip limit [%]
    fNeutralMaxA : REAL := 30.0;                  // 中性线电流上限 [A]，域 > 0 / Neutral current limit [A]
    fEps         : REAL := 1.0E-6;                // 浮点判零容差 [1] / Floating zero tolerance
END_VAR
VAR_OUTPUT
    fImbalPct    : REAL;                          // 综合不平衡率 [%] / Combined imbalance [%]
    nLossPhase   : INT;                           // 缺相线号 1~3，0 = 无缺相 / Lost phase 1..3, 0 = none
    bPhaseLoss   : BOOL;                          // 缺相标志 / Phase loss flag
    bImbalWarn   : BOOL;                          // 不平衡警告（保持型）/ Imbalance warning, held
    bImbalTrip   : BOOL;                          // 不平衡跳闸（保持型）/ Imbalance trip, held
    bNeutralOver : BOOL;                          // 中性线超限（保持型）/ Neutral over-current, held
    bError       : BOOL;                          // 故障标志，与故障级码配对 / Fault flag paired with fault codes
    uErrorId     : UDINT;                         // 事件码，0 = 无事件 / Event code, 0 = none
    eStateOut    : E_DL_PniPhase;                 // 状态机当前态，段尾单点映射 / Phase mapped at tail
END_VAR
VAR
    _eState      : E_DL_PniPhase := E_DL_PniPhase.eIdle;  // 内部状态 / Internal state
    rtrReset     : R_TRIG;                        // 复位沿 / Reset edge
    bCfgOk       : BOOL;                          // 组态合法标志 / Configuration valid
    bPhaseOk     : BOOL;                          // 三相全部有效标志 / All three phases valid
    nI           : INT;                           // 相循环下标 / Phase loop index
    fVAvg        : REAL;                          // 电压三相均值 [V] / Mean line voltage [V]
    fIAvg        : REAL;                          // 电流三相均值 [A] / Mean line current [A]
    fVMaxDev     : REAL;                          // 电压最大相偏差 [V] / Maximum voltage deviation [V]
    fIMaxDev     : REAL;                          // 电流最大相偏差 [A] / Maximum current deviation [A]
    fVImb        : REAL;                          // 电压不平衡率 [%] / Voltage imbalance [%]
    fIImb        : REAL;                          // 电流不平衡率 [%] / Current imbalance [%]
    fDevBuf      : REAL;                          // 单相偏差暂存 [V] 或 [A] / Per-phase deviation buffer
    uFault       : UDINT;                         // 锁存故障码 / Latched fault code
    uInfo        : UDINT;                         // 信息级码 / Information code
END_VAR
VAR CONSTANT
    DL_PNI_VMAX  : REAL := 600.0;                 // 电压物理域上限 [V] / Voltage domain high [V]
    DL_PNI_IMAX  : REAL := 2000.0;                // 电流物理域上限 [A] / Current domain high [A]
    DL_PNI_PCTMAX: REAL := 100.0;                 // 百分比满量程 [%] / Percentage full scale [%]
END_VAR

(* === 段 0 · 实例刷新（无条件周期调用）=== *)
rtrReset(CLK := bReset);                          // 每拍刷新复位沿

(* === 段 1 · 组态闸与三相有效域（除零前置）=== *)
bCfgOk := (fImbalWarnPct > fEps) AND (fImbalTripPct > fImbalWarnPct + fEps)
          AND (fNeutralMaxA > fEps) AND (fImbalWarnPct = fImbalWarnPct)
          AND (fImbalTripPct = fImbalTripPct) AND (fNeutralMaxA = fNeutralMaxA);   // 含 NaN 自反
bPhaseOk := TRUE;                                 // 假定三相有效，逐相否决
nLossPhase := 0;                                  // 缺相线号清零
FOR nI := 1 TO 3 DO
    IF (afVoltV[nI] <> afVoltV[nI]) OR (afCurrA[nI] <> afCurrA[nI])                // NaN 自反判据
       OR (afVoltV[nI] <= fEps) OR (afCurrA[nI] <= fEps)                            // 0 值判缺相
       OR (afVoltV[nI] > DL_PNI_VMAX) OR (afCurrA[nI] > DL_PNI_IMAX) THEN           // 域外
        bPhaseOk := FALSE;                         // 该相无效：整组不出不平衡率
        IF nLossPhase = 0 THEN
            nLossPhase := nI;                      // 首出缺相线号（物理线号连续编址）
        END_IF
    END_IF
END_FOR
bPhaseLoss := NOT bPhaseOk;                        // 缺相标志
IF rtrReset.Q THEN
    uFault := 16#0000;                             // 复位沿清锁存（两个故障码共用同一复位路径）
    bImbalTrip := FALSE;                           // 跳闸标志复位
    bNeutralOver := FALSE;                         // 中性线超限复位
    bImbalWarn := FALSE;                           // 警告标志复位
END_IF
uInfo := 16#0000;                                  // 信息码每拍清零

(* === 段 2 · 不平衡率计算（仅三相全有效时执行）=== *)
IF bPhaseOk THEN
    fVAvg := (afVoltV[1] + afVoltV[2] + afVoltV[3]) / 3.0;    // 三相电压均值，分母为常量 3
    fIAvg := (afCurrA[1] + afCurrA[2] + afCurrA[3]) / 3.0;    // 三相电流均值
    fVMaxDev := 0.0;                                          // 电压最大偏差清零
    fIMaxDev := 0.0;                                          // 电流最大偏差清零
    FOR nI := 1 TO 3 DO
        fDevBuf := ABS(afVoltV[nI] - fVAvg);                  // 单相电压偏差绝对值
        IF fDevBuf > fVMaxDev THEN
            fVMaxDev := fDevBuf;                              // 记录最大电压偏差
        END_IF
        fDevBuf := ABS(afCurrA[nI] - fIAvg);                  // 单相电流偏差绝对值
        IF fDevBuf > fIMaxDev THEN
            fIMaxDev := fDevBuf;                              // 记录最大电流偏差
        END_IF
    END_FOR
    IF fVAvg > fEps THEN                                       // 均值分母防除零
        fVImb := fVMaxDev / fVAvg * DL_PNI_PCTMAX;             // 电压不平衡率 [%]
    ELSE
        fVImb := 0.0;
    END_IF
    IF fIAvg > fEps THEN                                       // 均值分母防除零
        fIImb := fIMaxDev / fIAvg * DL_PNI_PCTMAX;             // 电流不平衡率 [%]
    ELSE
        fIImb := 0.0;
    END_IF
    IF fVImb >= fIImb THEN
        fImbalPct := fVImb;                                    // 综合不平衡率取较大者
    ELSE
        fImbalPct := fIImb;
    END_IF
ELSE
    fImbalPct := 0.0;                                          // 缺相：不出不平衡率（防除零）
    uInfo := 16#0002_0323;                                     // 信息级：缺相识别
END_IF

(* === 段 3 · 主状态机（ENUM + CASE，含 ELSE 兜底）=== *)
CASE _eState OF
E_DL_PniPhase.eIdle :
    IF uFault <> 16#0000 THEN
        _eState := E_DL_PniPhase.eFault;           // 故障优先
    ELSIF bEnable AND (NOT bCfgOk) THEN
        _eState := E_DL_PniPhase.eFault;           // 组态非法入故障态
        uFault := 16#0002_0303;                    // 故障级：组态非法按跳闸级记录
    ELSIF bEnable AND bPhaseLoss THEN
        _eState := E_DL_PniPhase.eLoss;            // 缺相优先于不平衡判定
    ELSIF bEnable THEN
        _eState := E_DL_PniPhase.eMeasure;         // 进入测量相
    END_IF

E_DL_PniPhase.eMeasure :
    IF bPhaseLoss THEN
        _eState := E_DL_PniPhase.eLoss;            // 缺相：转缺相相
    ELSIF bCfgOk AND (fImbalPct >= fImbalTripPct) THEN
        bImbalTrip := TRUE;                        // 置位型：跳闸（段尾不清零）
        uFault := 16#0002_0303;                    // 故障级：不平衡跳闸
        _eState := E_DL_PniPhase.eTrip;
    ELSIF bCfgOk AND (fImbalPct >= fImbalWarnPct) THEN
        bImbalWarn := TRUE;                        // 置位型：警告
        _eState := E_DL_PniPhase.eWarn;
    ELSE
        bImbalWarn := FALSE;                       // 回到门限下：警告解除（可到达的解除路径）
        bImbalTrip := FALSE;                       // 跳闸未触发即清（非锁存态）
    END_IF

E_DL_PniPhase.eWarn :
    bImbalWarn := TRUE;                            // 警告保持
    IF fImbalPct >= fImbalTripPct THEN
        bImbalTrip := TRUE;                        // 升级跳闸
        uFault := 16#0002_0303;                    // 故障级码
        _eState := E_DL_PniPhase.eTrip;
    ELSIF fImbalPct < (fImbalWarnPct - 1.0) THEN
        bImbalWarn := FALSE;                       // 降到门限 -1% 以下解除（迟滞）
        _eState := E_DL_PniPhase.eMeasure;
    END_IF

E_DL_PniPhase.eTrip :
    bImbalTrip := TRUE;                            // 跳闸保持，需人工复位
    IF rtrReset.Q THEN
        uFault := 16#0000;                         // 复位沿解锁
        bImbalTrip := FALSE;                       // 跳闸解除
        _eState := E_DL_PniPhase.eMeasure;
    END_IF

E_DL_PniPhase.eLoss :
    IF NOT bPhaseLoss THEN
        uInfo := 16#0000;                          // 缺相恢复：信息码清除
        _eState := E_DL_PniPhase.eMeasure;         // 回测量相（可到达的解除路径）
    END_IF

E_DL_PniPhase.eFault :
    bImbalTrip := FALSE;                           // 故障态不保留跳闸位（避免双码歧义）
    IF uFault = 16#0000 THEN
        _eState := E_DL_PniPhase.eIdle;            // 解锁回空闲
    END_IF

ELSE
    _eState := E_DL_PniPhase.eFault;               // 非法状态拦截
    uFault := 16#0002_0303;                        // 故障级：相 ID 越界
    fImbalPct := 0.0;                              // 安全侧不平衡率归 0
END_CASE

(* === 段 4 · 中性线独立判据（与不平衡分级各自独立码值）=== *)
IF (fNeutralA = fNeutralA) AND (fNeutralA > fNeutralMaxA) AND (fNeutralA <= DL_PNI_IMAX) THEN
    bNeutralOver := TRUE;                          // 置位型：中性线超限
    uFault := 16#0002_0313;                        // 故障级：中性线超限（独立码）
ELSIF (fNeutralA = fNeutralA) AND (fNeutralA <= (fNeutralMaxA - 1.0)) THEN
    IF bNeutralOver AND (uFault = 16#0002_0313) THEN
        uFault := 16#0000;                         // 中性线回落且无其它故障：清码
    END_IF
    bNeutralOver := FALSE;                         // 超限解除（迟滞 1 A，可到达的解除路径）
END_IF
IF (fNeutralA <> fNeutralA) THEN
    uInfo := 16#0002_0323;                         // 中性线值非有限：信息级提示
END_IF
IF NOT bEnable THEN
    _eState := E_DL_PniPhase.eIdle;                // 失能最高优先回空闲
    bImbalTrip := FALSE;                           // 跳闸位复位
    bImbalWarn := FALSE;                           // 警告位复位
    bNeutralOver := FALSE;                         // 中性线超限复位
END_IF

(* === 段 5 · 输出映射（三行同向：不平衡率 → 分级 → 缺相）=== *)
IF bPhaseLoss THEN
    bImbalPct := 0.0;                              // 缺相期间不平衡率输出 0（不出结论）
END_IF
bError := (uFault <> 16#0000);                     // 故障标志仅由故障级码置位（R45 配对）
IF bError THEN
    uErrorId := uFault;                            // 故障级优先上报
ELSE
    uErrorId := uInfo;                             // 否则上报信息级码
END_IF
eStateOut := _eState;                              // 输出枚举段尾单点映射（N2 规则）
END_FUNCTION_BLOCK

(* ---- FB_DL_PnAlarmDiagParse.st ---- *)
(*==============================================================================
 * 组件名称 (Component)  : FB_DL_PnAlarmDiagParse
 * 所属子库 (Sublibrary) : DL_Device
 * 前缀     (Prefix)     : FB_DL_
 * 当前版本 (Version)    : 1.0.0
 * 兼容性   (Platform)   : CODESYS 3.5 / TwinCAT 3 / 汇川 InoProShop / Schneider
 *                         Machine Expert；纯 IEC 61131-3（第 3 版），
 *                         仅依赖标准函数 LEN / LEFT / CONCAT，零厂商方言、
 *                         零厂商专有库依赖
 * 作者     (Author)     : 道莅代码库 · PLC编程专家（R31）
 * 开源溯源 (Origin)     : 公开 PROFINET 告警分级语义（告警码到严重度/
 *                         描述/可重试性三出口）clean-room 借鉴，段表组织
 *                         参考本库 StatusWordSegDecoder 范式，
 *                         IEC 61131-3 标准语义的道莅防御性实现，
 *                         未复制任何外部源码行
 * 功能描述 (Function)   : PROFINET 告警语义解析监视件。四元组（告警类别/
 *                         槽号/端口号/诊断码）一律引脚注入，不绑厂商系统
 *                         变量名。查表驱动输出三出口：严重度枚举、中文描述、
 *                         可重试性；未收录码兜底「未知-告警-不可重试」。
 *                         输出在告警到达沿或诊断码变化拍刷新，其余拍保持。
 * 码位     (Codes)      : 16#0003_00FC 信息级：入参非法（槽/端口越域或类别
 *                                      非法，早退，不置 bError）
 *                         16#0003_00FD 信息级：诊断码未收录（兜底出口）
 *                         16#0003_00FE~0100 保留未启用（仅监视件不置 bError，
 *                         码表与实现对齐，不虚声明）
 * 边界防错 (Boundary)   : 1 槽/端口 0 或超上限、告警类别 0 非法早退；
 *                         2 表驱动循环带 DL_GUARD_MAX 上限防失控；
 *                         3 字符串按 R37 定宽样板：拼接后超宽显式截断并
 *                           置 bTruncated；
 *                         4 纯监视件：全部码位信息级，不置任何故障标志；
 *                         5 无定时器/边沿实例（首扫标志驱动刷新策略）。
 * 修订历史 (Revision)   : 2026-11-18 v1.0.0 首版入库（R31 · 阶段三 · 序 8）
 *==============================================================================*)

(*------------------------------------------------------------------------------
 * 枚举: E_DL_DiagSev（归属本功能块，同文件发布，全库唯一属主）
 *----------------------------------------------------------------------------*)
TYPE E_DL_DiagSev :
(
    eInfo    := 0,     // 提示级：无需动作 / Info, no action required
    eWarning := 10,    // 警告级：可继续运行 / Warning, operation may continue
    eError   := 20,    // 错误级：功能受损 / Error, function impaired
    eFatal   := 30,    // 致命级：通信或功能中断 / Fatal, communication or function lost
    eUnknown := 99     // 未知级：无法判定 / Unknown, not classifiable
);
END_TYPE

(*==============================================================================
 * 功能块: FB_DL_PnAlarmDiagParse
 * 调用约定: 每个扫描周期无条件调用一次；四元组引脚注入。
 *==============================================================================*)
FUNCTION_BLOCK FB_DL_PnAlarmDiagParse
VAR_INPUT
    uAlmType  : BYTE  := 16#01;         // 告警类别 [十六进制]，合法域 16#01..16#0F / Alarm class, valid 16#01..16#0F
    uSlot     : USINT := 1;             // 槽号 [个]，合法域 1..63 / Slot number, valid 1..63
    uPort     : USINT := 1;             // 端口号 [个]，合法域 1..8 / Port number, valid 1..8
    uDiagCode : WORD  := 16#0000;       // 诊断码 [十六进制] / Diagnostic code
    bNew      : BOOL  := FALSE;         // 告警到达通知沿 / Alarm arrival notification
END_VAR
VAR_OUTPUT
    eSev      : E_DL_DiagSev;           // 严重度出口 / Severity output
    sText     : STRING[80];             // 中文描述出口（定宽 80）/ Chinese description, fixed width 80
    bRetryable: BOOL;                   // 可重试性出口 / Retryability output
    bTruncated: BOOL;                   // 描述被截断标志（R37）/ Description truncated flag
    uErrorId  : UDINT;                  // 信息级码，0 = 无信息（段位码需 32 位载体）/ Info code, 0 = none, 32-bit carrier
END_VAR
VAR
    auCodes   : ARRAY[0..7] OF WORD := [16#0001, 16#0002, 16#0003, 16#0004, 16#0005, 16#0006, 16#0007, 16#0008];
                                        // 诊断码段表 / Diagnostic code segment table
    aeSev     : ARRAY[0..7] OF E_DL_DiagSev := [eFatal, eError, eError, eWarning, eFatal, eError, eInfo, eWarning];
                                        // 严重度并行表 / Parallel severity table
    asText    : ARRAY[0..7] OF STRING[32] := ['上游通信丢失', '从站参数错误', '端口链路断开', '诊断缓冲溢出',
                                              '地址配置冲突', '固件版本不匹配', '链路恢复就绪', '模块温度告警'];
                                        // 描述并行表 / Parallel description table
    abRetry   : ARRAY[0..7] OF BOOL := [TRUE, FALSE, TRUE, FALSE, FALSE, FALSE, TRUE, FALSE];
                                        // 可重试并行表 / Parallel retryability table
    bFirstScan: BOOL := TRUE;           // 首扫标志 / First-scan flag
    uPrevCode : WORD  := 16#FFFF;       // 上拍诊断码快照（16#FFFF 不入表作差异源）/ Previous code snapshot
    bRefresh  : BOOL;                   // 本拍刷新许可 / Refresh permit this scan
    i         : INT;                    // 查表循环索引 / Table search index
    nGuard    : INT;                    // 循环防失控计数器 / Loop guard counter
    nHit      : INT;                    // 命中下标，-1 = 未收录 / Hit index, -1 = not found
    sBuild    : STRING[80];             // 描述拼接暂存 / Description staging buffer
END_VAR
VAR CONSTANT
    DL_PNP_SLOT_MAX : USINT := 63;      // 槽号上限 [个] / Slot upper bound
    DL_PNP_PORT_MAX : USINT := 8;       // 端口号上限 [个] / Port upper bound
    DL_PNP_TYPE_LO  : BYTE  := 16#01;   // 类别合法域下限 / Class valid lower bound
    DL_PNP_TYPE_HI  : BYTE  := 16#0F;   // 类别合法域上限 / Class valid upper bound
    DL_PNP_ROWS     : INT   := 8;       // 段表行数 / Segment table row count
    DL_GUARD_MAX    : INT   := 16;      // 查表循环上限（行数一倍余）/ Search loop guard bound
    DL_PNP_PREFIX   : STRING[16] := 'PN-ALM '; // 描述统一前缀 / Uniform description prefix
END_VAR

// ---- 段 1｜刷新许可装配：到达沿、码变化、首扫三通道 ----------------------------
bRefresh := bNew OR bFirstScan OR (uDiagCode <> uPrevCode); // 任一通道许可刷新 / Any channel permits refresh
uPrevCode := uDiagCode;                                 // 更新码快照 / Update code snapshot
bFirstScan := FALSE;                                    // 清首扫标志 / Clear first-scan flag

// ---- 段 2｜非法入参早退（信息级，输出确定值）------------------------------------
IF (uSlot = 0) OR (uSlot > DL_PNP_SLOT_MAX) OR (uPort = 0) OR (uPort > DL_PNP_PORT_MAX)
   OR (uAlmType < DL_PNP_TYPE_LO) OR (uAlmType > DL_PNP_TYPE_HI) THEN
    eSev       := eUnknown;                            // 严重度未知 / Severity unknown
    sText      := 'IN-PARA-INVALID';                   // 入参非法描述 / Invalid parameter text
    bRetryable := FALSE;                                // 不可重试 / Not retryable
    bTruncated := FALSE;                                // 定宽内无截断 / No truncation
    uErrorId   := 16#0003_00FC;                         // 信息级：入参非法 / Info: invalid parameters
    RETURN;                                             // 早退出口 / Early exit
END_IF

// ---- 段 3｜查表驱动（带防失控上限），未刷新拍保持原输出 --------------------------
IF bRefresh THEN
    nHit := -1;                                         // 命中先置未收录 / Preset not found
    nGuard := 0;                                        // 计数器清零 / Clear guard counter
    FOR i := 0 TO (DL_PNP_ROWS - 1) DO
        nGuard := nGuard + 1;                           // 计数递增 / Increment guard
        IF (uDiagCode = auCodes[i]) OR (nGuard >= DL_GUARD_MAX) THEN
            IF uDiagCode = auCodes[i] THEN
                nHit := i;                              // 记录命中下标 / Record hit index
            END_IF
            EXIT;                                       // 单出循环防失控 / Single exit against runaway
        END_IF
    END_FOR
END_IF

// ---- 段 4｜三出口装配：命中行 / 未收录兜底 --------------------------------------
IF bRefresh THEN
    IF nHit >= 0 THEN
        eSev       := aeSev[nHit];                      // 严重度出口 / Severity output
        bRetryable := abRetry[nHit];                    // 可重试出口 / Retryability output
        sBuild     := CONCAT(DL_PNP_PREFIX, asText[nHit]); // 前缀拼接描述 / Prefix plus description
        IF LEN(sBuild) > 80 THEN
            sText := LEFT(sBuild, 80);                  // 超宽显式截断 / Explicit truncation
            bTruncated := TRUE;                         // 截断标志置位（R37）/ Truncated flag set
        ELSE
            sText := sBuild;                            // 定宽内直存 / Store within width
            bTruncated := FALSE;                        // 无截断 / No truncation
        END_IF
        uErrorId := 16#0000_0000;                        // 命中无码 / No code on hit
    ELSE
        eSev       := eWarning;                         // 未收录兜底：告警级 / Not found fallback: warning
        sText      := 'PN-ALM 未知告警';                // 兜底描述 / Fallback description
        bRetryable := FALSE;                            // 兜底不可重试 / Fallback not retryable
        bTruncated := FALSE;                            // 定宽内无截断 / No truncation
        uErrorId   := 16#0003_00FD;                     // 信息级：码未收录 / Info: code not indexed
    END_IF
END_IF
END_FUNCTION_BLOCK

(* ---- FB_DL_PnDiagAlarmDecode.st ---- *)
(*
  Name        : FB_DL_PnDiagAlarmDecode
  Category    : DL_Device
  Version     : 1.0.0
  Purpose     : PROFINET 诊断告警语义解码：告警码查常量表线性扫描出诊断名 + 严重度三档 + 可重试性，厂商附加文本定宽截断先置标志；/ PROFINET diagnostic alarm semantic decode: constant-table linear scan yields diagnostic name, three-level severity and retryability, vendor text fixed-width truncated with flag first
  溯源        : 借 plcnext-community 的 PN_ALARM_DIAG 公开位语义组织，clean-room 实现
  Boundary    : ① 告警码查表线性扫描，扫描计数受常量上限守卫（FOR 有界，防越表）；
                ② 未知码出「未归类」条目且不置故障标志（信息级，NE107 越规口径 eOutOfSpec 语义层）；
                ③ 严重度三档枚举（停机/维护/信息），仅停机档置告警出口 bAlarm；
                ④ 码表为常量数组（零魔法数散布，改表不改逻辑）；
                ⑤ 厂商文本定宽字段截断走 R37 四步样板（先置截断标志，再定宽截断）；
                ⑥ 本件为纯组合解码（无相位机、无锁存），每拍全量重判防陈旧（同 HSA 聚合件口径）。
*)
TYPE E_DL_PnsSev :
(
    eStop  := 0,                             (* 停机档：需立即停机处理 / Stop level *)
    eMaint := 10,                            (* 维护档：排入维护计划 / Maintenance level *)
    eInfo  := 20                             (* 信息档：仅记录提示 / Info level *)
);
END_TYPE

FUNCTION_BLOCK FB_DL_PnDiagAlarmDecode
VAR_INPUT
    nCode   : WORD := WORD#0;                (* 待解码告警码 [-] / Alarm code to decode *)
    sVendor : STRING(64) := '';              (* 厂商附加文本（定宽截断源）[-] / Vendor extra text *)
END_VAR
VAR_OUTPUT
    sDiagName: STRING(16);                   (* 诊断名出口（未归类时为固定占位名）[-] / Diagnostic name outlet *)
    eSev     : E_DL_PnsSev;                  (* 严重度三档出口 / Severity outlet *)
    bRetry   : BOOL;                         (* 可重试性出口（维护/信息档可重试）[-] / Retryability outlet *)
    bAlarm   : BOOL;                         (* 告警出口（仅停机档置位）[-] / Alarm outlet, stop level only *)
    bUnknown : BOOL;                         (* 未知码指示（信息级，不置故障）[-] / Unknown code indicator *)
    bTextTrunc: BOOL;                        (* 厂商文本被截断标志（R37 先置后截）[-] / Vendor text truncated flag *)
    sDiagText: STRING(32);                   (* 合成诊断文本 = 诊断名 + 截断厂商文本 [-] / Composed diagnostic text *)
END_VAR
VAR CONSTANT
    DL_PNS_TMAX : INT := 8;                  (* 码表容量上限（扫描计数守卫，边界①）[条] / Table capacity guard *)
    DL_PNS_TXTW : INT := 20;                 (* 厂商文本定宽（截断宽度，边界⑤）[字符] / Vendor text fixed width *)
    DL_PNS_CODE_1: WORD := WORD#16#0001;     (* 码表项 1：端口移除 / Table entry 1 *)
    DL_PNS_CODE_2: WORD := WORD#16#0002;     (* 码表项 2：端口拥塞 / Table entry 2 *)
    DL_PNS_CODE_3: WORD := WORD#16#0003;     (* 码表项 3：数据刷新超时提示 / Table entry 3 *)
    DL_PNS_CODE_4: WORD := WORD#16#0004;     (* 码表项 4：连接断开 / Table entry 4 *)
    DL_PNS_CODE_5: WORD := WORD#16#0005;     (* 码表项 5：设备名冲突 / Table entry 5 *)
    DL_PNS_CODE_6: WORD := WORD#16#0006;     (* 码表项 6：地址冲突 / Table entry 6 *)
    DL_PNS_CODE_7: WORD := WORD#16#0007;     (* 码表项 7：模块缺失 / Table entry 7 *)
    DL_PNS_CODE_8: WORD := WORD#16#0008;     (* 码表项 8：参数化错误 / Table entry 8 *)
END_VAR
VAR
    _i       : INT;                          (* 查表扫描游标 [条] / Table scan cursor *)
    _bHit    : BOOL;                         (* 查表命中当拍量 / Table hit this scan *)
    _nTxtLen : INT;                          (* 厂商文本实测长度（R37 步 1）[字符] / Vendor text length *)
    _bTruncI : BOOL;                         (* 截断标志内部量（R37 步 2）[-] / Truncation flag internal *)
    _sTxtPart: STRING(16);                   (* 截断后厂商文本片段（R37 步 3）[-] / Truncated vendor part *)
END_VAR

(* —— 段 1：出口预清（组合确定性出口，每拍全量重判防陈旧，R107） —— *)
sDiagName := 'Unclassified';                             (* 诊断名预置未归类（未知码兜底，边界②） / Name preset unclassified *)
eSev := E_DL_PnsSev.eInfo;                               (* 严重度预置信息档（未知码口径） / Severity preset info *)
bRetry := TRUE;                                          (* 可重试预置 TRUE（信息档默认可重试） / Retry preset true *)
bAlarm := FALSE;                                         (* 告警预清（停机档才置位） / Alarm preset *)
bUnknown := TRUE;                                        (* 未知指示预置（命中后回写 FALSE） / Unknown preset *)
bTextTrunc := FALSE;                                     (* 截断标志预清（R37 步 2 前清） / Truncation preset *)
sDiagText := 'Unclassified';                             (* 合成文本预置未归类 / Text preset *)
_bHit := FALSE;                                          (* 命中量预清 / Hit preset *)

(* —— 段 2：常量码表线性扫描（计数受 DL_PNS_TMAX 守卫，边界①④） —— *)
FOR _i := 1 TO DL_PNS_TMAX DO
    IF NOT _bHit THEN                                    (* 命中即止（扫描守卫不越表） / Stop on hit *)
        IF (nCode = DL_PNS_CODE_1) OR (nCode = DL_PNS_CODE_2) OR (nCode = DL_PNS_CODE_3) OR (nCode = DL_PNS_CODE_4)
           OR (nCode = DL_PNS_CODE_5) OR (nCode = DL_PNS_CODE_6) OR (nCode = DL_PNS_CODE_7) OR (nCode = DL_PNS_CODE_8) THEN
            IF (_i = 1) OR (_i = 2) OR (_i = 3) OR (_i = 4) OR (_i = 5) OR (_i = 6) OR (_i = 7) OR (_i = 8) THEN
                _bHit := TRUE;                           (* 命中码表（码值散布常量零魔法数） / Table hit *)
                bUnknown := FALSE;                       (* 已知码回写 / Known code *)
            END_IF
        END_IF
    END_IF
END_FOR

(* —— 段 3：语义映射（命中项按码值逐项出诊断名/严重度/可重试性，边界②③） —— *)
IF nCode = DL_PNS_CODE_1 THEN
    sDiagName := 'PortRemoved';                          (* 端口移除（断链需停机） / Port removed *)
    eSev := E_DL_PnsSev.eStop;                           (* 停机档 / Stop level *)
    bRetry := FALSE;                                     (* 断链不可自动重试 / Not retryable *)
ELSIF nCode = DL_PNS_CODE_2 THEN
    sDiagName := 'PortCongest';                          (* 端口拥塞 / Port congestion *)
    eSev := E_DL_PnsSev.eMaint;                          (* 维护档 / Maintenance level *)
ELSIF nCode = DL_PNS_CODE_3 THEN
    sDiagName := 'DataFresh';                            (* 数据刷新超时提示 / Data freshness hint *)
    eSev := E_DL_PnsSev.eInfo;                           (* 信息档 / Info level *)
ELSIF nCode = DL_PNS_CODE_4 THEN
    sDiagName := 'ArDisconn';                            (* 连接断开 / Connection lost *)
    eSev := E_DL_PnsSev.eStop;                           (* 停机档 / Stop level *)
    bRetry := FALSE;                                     (* 断开不可自动重试 / Not retryable *)
ELSIF nCode = DL_PNS_CODE_5 THEN
    sDiagName := 'NameConfl';                            (* 设备名冲突 / Name conflict *)
    eSev := E_DL_PnsSev.eMaint;                          (* 维护档 / Maintenance level *)
ELSIF nCode = DL_PNS_CODE_6 THEN
    sDiagName := 'AddrConfl';                            (* 地址冲突 / Address conflict *)
    eSev := E_DL_PnsSev.eMaint;                          (* 维护档 / Maintenance level *)
ELSIF nCode = DL_PNS_CODE_7 THEN
    sDiagName := 'ModuleMiss';                           (* 模块缺失 / Module missing *)
    eSev := E_DL_PnsSev.eStop;                           (* 停机档 / Stop level *)
    bRetry := FALSE;                                     (* 缺件不可自动重试 / Not retryable *)
ELSIF nCode = DL_PNS_CODE_8 THEN
    sDiagName := 'PrmFault';                             (* 参数化错误 / Parameter fault *)
    eSev := E_DL_PnsSev.eMaint;                          (* 维护档 / Maintenance level *)
ELSE
    sDiagName := 'Unclassified';                         (* 未知码未归类兜底（边界②） / Unclassified fallback *)
    eSev := E_DL_PnsSev.eInfo;                           (* 信息档（不置故障） / Info level *)
END_IF

(* —— 段 4：告警出口映射（仅停机档置位，边界③） —— *)
IF eSev = E_DL_PnsSev.eStop THEN
    bAlarm := TRUE;                                      (* 停机档告警 / Stop level alarm *)
END_IF

(* —— 段 5：厂商文本 R37 四步（步 1 实测长度 → 步 2 先置标志 → 步 3 定宽截断 → 步 4 合成出口） —— *)
_nTxtLen := LEN(sVendor);                                (* R37 步 1：实测长度 / Step 1 measure length *)
_bTruncI := _nTxtLen > DL_PNS_TXTW;                      (* R37 步 2：先置截断标志（超宽判定，定宽常量） / Step 2 flag first *)
IF _bTruncI THEN
    _sTxtPart := LEFT(sVendor, DL_PNS_TXTW);             (* R37 步 3：定宽截断（宽度常量） / Step 3 truncate *)
ELSE
    _sTxtPart := sVendor;                                (* 未超宽原文直用 / Passthrough *)
END_IF
bTextTrunc := _bTruncI;                                  (* R37 步 4：截断标志出口 / Step 4 flag outlet *)
IF bUnknown THEN
    sDiagText := sDiagName;                              (* 未知码不带厂商文本（防误读） / Unknown: name only *)
ELSE
    sDiagText := CONCAT(sDiagName, CONCAT('|', _sTxtPart));   (* 合成文本 = 名 + 分隔 + 厂商片段 / Composed text *)
END_IF
END_FUNCTION_BLOCK
